(* IEC 61131-3 sources: daoli-st-library/DL_MathData (part 19) *)

(* ---- FC_DL_MeanAbsDevCalc.st ---- *)
(*
  ==================================================================
  组件名 Component  : FC_DL_MeanAbsDevCalc
  分类   Category   : DL_MathData
  前缀   Naming     : FC_DL_ ｜ b/n/u/f/t/e/st 类型前缀制（R265）
  复杂度 Complexity  : 低
  版本   Version    : 1.0.0
  功能   Purpose    : 均值绝对偏差 MAD-mean = mean(|xᵢ − mean|)，两遍法。
  来源   Source     : self-std（公开统计语义自研）
  平台   Platform   : 纯 IEC 61131-3（FOR / 四则 / ABS），三平台通用
  分工声明 Split     : 与 FC_DL_MedianAbsDev（中位数域属主）分工——后者以中位数
                      为中心（对离群点稳健）；本件以均值为中心（R216 双向互引）。
  作者   Author     : 道莅代码库 · PLC 编程专家（R61）
  归属 Ownership     : 本件无 TYPE 声明；引用件类型全部 IEC 标准原生。
  ------------------------------------------------------------------
  边界 Boundary     :
                      一 nCount < 1 置信息级码不计算（nCount = 0 无均值可言）；
                      二 计数 > 256 钳位续算置信息级；
                      三 元素非有限逐个点名判故障拒绝（R272 全量）；
                      四 均值非有限传播闸：均值算出后复检，非有限同判故障；
                      五 除子 nUse 已证 ≥ 1（域闸下界），无除零风险；
                      六 结果复检兜底同拍置 eErr + bError + bValid 三件套（R258）；
                      七 只读入参数组，不改调用方数据；无状态纯函数（R254）。
  错误码   Codes    :
    16#0001_063C【信息级】计数越域已钳位（<1 早退，>256 钳位续算）
    16#0001_063D【故障级】元素或均值非有限，拒绝出值
  验收   Acceptance :
    算法已证（脚本）：未跑 ｜ 编译器已证（三平台）：未跑
    V1 值 1/2/3 → mean=2、MAD-mean=2/3；V2 值 5/5/5 → 0
    V3 nCount=0 → 码 063C、bValid=FALSE；V4 含 NaN → 码 063D、bError=TRUE
  修订记录 Revision  :
    2026-11-21  v1.0.0  R61 首版（批 2 · 序号 7）
  ==================================================================
*)
FUNCTION FC_DL_MeanAbsDevCalc : BOOL
VAR_IN_OUT
    afValues : ARRAY[0..255] OF LREAL; // 数值序列 [工程单位]，只读 / the value series, read only
END_VAR
VAR_INPUT
    nCount : DINT; // 序列个数 [个]，合法域 1..256 / the count, legal from one to two hundred fifty six
END_VAR
VAR_OUTPUT
    fMad   : LREAL; // 均值绝对偏差 [工程单位] / the mean absolute deviation
    fMean  : LREAL; // 序列均值 [工程单位] / the series mean
    bValid : BOOL;  // 结果可用标志 [-] / the result usable flag
    eErr   : UDINT; // 错误码，0 = 正常 / the error code, zero is ok
    bError : BOOL;  // 错误标志，故障级码置位（R45 配对）/ the error flag
END_VAR
VAR
    k     : DINT;  // 遍历索引 [下标] / the traversal index
    nUse  : DINT;  // 钳位后的个数 [个] / the clamped count
    fSum  : LREAL; // 一遍和累加器 [工程单位] / the first pass sum accumulator
    fDev  : LREAL; // 二遍偏差累加器 [工程单位] / the second pass deviation accumulator
END_VAR
VAR CONSTANT
    DL_MAD_NMAX : DINT := 256; // 序列容量上界 [个]，与数组容量一致 / the capacity aligned with the array
END_VAR

// 段 1｜返回值与错误状态预置安全值 + 局部量显式预置（R45 / R254）/ segment 1, the preset
FC_DL_MeanAbsDevCalc := FALSE; // 返回值预置假 / preset the return false
fMad := 0.0; // 偏差预置零 / preset the deviation zero
fMean := 0.0; // 均值预置零 / preset the mean zero
bValid := FALSE; // 有效标志预置假 / preset the validity false
eErr := 16#0000_0000; // 错误码预置正常 / preset the code to ok
bError := FALSE; // 错误标志预置假 / preset the error flag false
nUse := 0; // 个数预置零 / preset the count zero
fSum := 0.0; // 一遍和预置零 / preset the sum zero
fDev := 0.0; // 二遍偏差预置零 / preset the deviation accumulator zero

// 段 2｜计数域闸（<1 早退，>256 钳位，边界一二）/ segment 2, the count gate
IF nCount < 1 THEN // 空序列无均值（边界一）/ an empty series has no mean
    eErr := 16#0001_063C; // 信息级：计数越域已钳位（信息级不置 bError）/ informational, the count clamped
    RETURN; // 早退 / early return
END_IF
nUse := nCount; // 域内接管 / take the count
IF nUse > DL_MAD_NMAX THEN // 超容量（边界二）/ above the capacity
    nUse := DL_MAD_NMAX; // 钳到容量 / clamp to the capacity
    eErr := 16#0001_063C; // 信息级：计数越域已钳位 / informational, the count clamped
END_IF

// 段 3｜一遍求和 + 元素非有限逐个点名（R272，边界三）/ segment 3, the first pass sum with the element wise gate
FOR k := 0 TO nUse - 1 DO // 有界遍历 / the bounded traversal
    IF (afValues[k] <> afValues[k]) OR ((afValues[k] - afValues[k]) <> (afValues[k] - afValues[k])) THEN // 元素非有限 / the element is not finite
        eErr := 16#0001_063D; // 故障级：元素非有限 / fault grade, a non finite element
        bError := TRUE; // 置错误标志（R45 配对）/ raise the error flag
        RETURN; // 早退 / early return
    END_IF
    fSum := fSum + afValues[k]; // 求和累加 / accumulate the sum
END_FOR
fMean := fSum / DINT_TO_LREAL(nUse); // 均值（除子已证 ≥ 1，边界五）/ the mean with a proven divisor
IF (fMean <> fMean) OR ((fMean - fMean) <> (fMean - fMean)) THEN // 均值非有限传播闸（边界四）/ the mean finiteness gate
    eErr := 16#0001_063D; // 故障级：均值非有限 / fault grade, a non finite mean
    bError := TRUE; // 置错误标志（R45 配对）/ raise the error flag
    RETURN; // 早退 / early return
END_IF

// 段 4｜二遍偏差累加（均值已证有限）/ segment 4, the second pass deviation accumulation
FOR k := 0 TO nUse - 1 DO // 有界遍历 / the bounded traversal
    fDev := fDev + ABS(afValues[k] - fMean); // 绝对偏差累加 / accumulate the absolute deviation
END_FOR
fMad := fDev / DINT_TO_LREAL(nUse); // 偏差均值（除子 nUse 已证 ≥ 1，同段 3 口径）/ the deviation mean with the proven divisor

// 段 5｜结果复检兜底（非有限同拍三件套，边界六）/ segment 5, the result recheck
IF (fMad <> fMad) OR ((fMad - fMad) <> (fMad - fMad)) THEN // 结果非有限 / the result is not finite
    fMad := 0.0; // 兜底安全值 / the bottom line safe value
    eErr := 16#0001_063D; // 故障级：结果非有限 / fault grade, the non finite result
    bError := TRUE; // 置错误标志（R45 配对）/ raise the error flag
    bValid := FALSE; // 结果不可用 / the result void
    RETURN; // 早退 / early return
END_IF
bValid := TRUE; // 结果可用 / the result is usable
FC_DL_MeanAbsDevCalc := TRUE; // 返回成功 / return success
END_FUNCTION

(* ---- FC_DL_MedianAbsDev.st ---- *)
(*==============================================================================
 * 组件名称 (Component)  : FC_DL_MedianAbsDev
 * 所属子库 (Sublibrary) : DL_MathData
 * 当前版本 (Version)    : 1.0.0
 * 兼容性   (Platform)   : CODESYS 3.5+ / TwinCAT 3 / 汇川 InoProShop / 施耐德 Machine Expert
 *                         仅用 FOR 循环、赋值与 ABS，无任何厂商内建函数（连排序库都不用）
 * 功能描述 (Function)   : 中位绝对偏差 MAD（Median Absolute Deviation），鲁棒离散度指标。
 *                           步骤：① 取前 nCount 个样本复制到本地缓冲（不改调用方数组）；
 *                                 ② 插入排序求中位数 fMedian；
 *                                 ③ 各样本减中位数取绝对值，再次插入排序求中位数 fMad。
 *                         返回 fMad。MAD 对离群点不敏感（崩溃点 50%），在传感器脏数据、
 *                         偶发尖峰场景下比标准差可靠：一个 10 倍离群点能把标准差抬高数倍，
 *                         而 MAD 几乎不变。
 *                         小样本策略：nCount < 3 → 无稳健意义，bValid=FALSE、返回 0；
 *                         nCount > 16 → 钳到 16（缓冲上界），bClamped=TRUE，结果按前 16 个算。
 *                         偶数样本的中位数取中间两数的算术平均（IEC 惯例，写死在此）。
 * 无状态边界 (Stateless): **本 FC 零内部状态**——本地缓冲 afWork / afDev 均为 VAR 临时量，
 *                         每次调用重新填装；IEC 61131-3 的 FC 本就不允许持有静态变量，本件遵守。
 *                         因此同一组样本重复调用结果完全一致，可重入、可并发、可放在任意 POU。
 *                         调用方若需"跨窗统计"，请自行保存样本数组，而不是期望 FC 记住上次数据。
 * 接口     (Interface)  : 入 afSample 样本数组（VAR_IN_OUT，本件只读，按 nCount 截取）、
 *                         nCount 有效样本数（1..16）；出 fMedian 中位数、fMad 中位绝对偏差、
 *                         bValid 结果有效（nCount >= 3）、bClamped 样本数被钳到 16。
 * 边界     (Boundary)   : ① 样本数下限：nCount < 3 无稳健离散意义 → bValid=FALSE、fMedian/fMad 置 0
 *                         （**0 不是"无离散"的断言**，调用方须查 bValid）；
 *                         ② 样本数上限：nCount > 16 → 钳到 16 并置 bClamped（绝不越 ARRAY 上界）；
 *                         ③ nCount <= 0 → bValid=FALSE、返回 0（防 nCount−1 为负导致的循环越界）；
 *                         ④ 非有限样本（NaN/Inf）会让排序结果失去意义：本件**不静默吞掉**，
 *                         检出即 bNonFin=TRUE、bValid=FALSE、返回 0（宁可不报，不可乱报）；
 *                         ⑤ 插入排序 O(n²)，n<=16 时最坏 256 次比较/两轮，代价可接受且无递归。
 * 依赖     (Depends)    : 无 DL_ 内部依赖；无标准库功能块依赖
 * 来源标签 (Source Tag) : T2-1 ◐（MAD 为公开经典鲁棒统计量，Hampel 1974；插入排序为教科书算法；
 *                         ST 实现为道莅自研，零代码行复制）
 * 码表     (Codes)      : 本件不占用任何全局数字码位。异常出口为 BOOL（bValid / bClamped / bNonFin）；
 *                         数字码位待主控收口阶段统一派号。
 * 红线自检 (Redline)    : R1 ✓ 零 GVL/VAR_EXTERNAL ｜ R2 ✓ 零 %I/%Q/%M ｜ R3 ✓ 纯 IEC 61131-3
 *                         R4 ✓ 数组边界钳位 + 循环上界由钳位量派生 + 非有限闸
 *                         R5 ✓ 声明逐行同行双语注释 ｜ R6 N/A（无状态机）
 *                         R7 N/A（无实例调用）
 * 修订历史 (Revision)   : 2026-11-19  v1.0.0  R46 首版（批次 3 · 序号 15）
 *==============================================================================*)
FUNCTION FC_DL_MedianAbsDev : REAL
VAR_IN_OUT
    afSample : ARRAY[0..15] OF REAL;    // 样本数组（本件只读，按 nCount 截取） [工程单位] / Sample array, read-only here, sliced by nCount
END_VAR
VAR_INPUT
    nCount : INT := 3;                  // 有效样本数，域 1..16（>16 被钳位） [个] / Valid sample count, 1..16, clamped above
END_VAR
VAR_OUTPUT
    fMedian  : REAL;                    // 样本中位数 [工程单位] / Sample median [engineering unit]
    bValid   : BOOL;                    // 结果有效（3 <= 有效样本数 <= 16） [-] / Result valid
    bClamped : BOOL;                    // 样本数被钳到 16 [-] / Sample count clamped to 16
    bNonFin  : BOOL;                    // 样本中存在 NaN/Inf，结果不可信 [-] / A non-finite sample was found
END_VAR
VAR
    afWork : ARRAY[0..15] OF REAL;      // 工作副本（排序用，不动调用方数组） [工程单位] / Working copy for sorting
    afDev  : ARRAY[0..15] OF REAL;      // 绝对偏差数组（排序用） [工程单位] / Absolute-deviation array for sorting
    nUse   : INT;                       // 实际参与计算的样本数（钳位后） [个] / Actual sample count after clamping
    i      : INT;                       // 外层遍历索引 / Outer loop index
    j      : INT;                       // 插入排序内层索引 / Inner index for the insertion sort
    fKey   : REAL;                      // 插入排序暂存键 [工程单位] / Key kept while inserting
    fLo    : REAL;                      // 偶数样本时中位数取中间两值之一 [工程单位] / One of the two middle values
    fHi    : REAL;                      // 偶数样本时中位数取中间两值之另一 [工程单位] / The other middle value
    nMidi  : INT;                       // 中位数取位下标（下中位） [个] / Lower middle index
END_VAR
VAR CONSTANT
    DL_MAD_MAXN : INT := 16;            // 样本容量（与 ARRAY 上界一致） [个] / Sample capacity matching the array bounds
    DL_MAD_MINN : INT := 3;             // 稳健统计所需最少样本数 [个] / Minimum sample count for robust statistics
END_VAR

(* —— 段 1：出口初始化（任何路径下返回值确定） —— *)
FC_DL_MedianAbsDev := 0.0;      // 缺省返回 0，须配 bValid 才可用 / Default 0, meaningful only with bValid
fMedian  := 0.0;                // 中位数清零 / Median cleared
bValid   := FALSE;              // 先假定无效 / Assume invalid
bClamped := FALSE;              // 钳位标志清零 / Clamp flag cleared
bNonFin  := FALSE;              // 非有限标志清零 / Non-finite flag cleared

(* —— 段 2：样本数钳位（先钳后循环，循环上界全部由 nUse 派生） —— *)
IF nCount <= 0 THEN
    RETURN;                     // 无样本：直接返回哨兵 0 / No samples: return the sentinel
END_IF
nUse := nCount;                 // 取请求样本数 / Take the requested count
IF nUse > DL_MAD_MAXN THEN
    nUse := DL_MAD_MAXN;        // 上界钳到容量 / Clamp to capacity
    bClamped := TRUE;           // 标记被钳 / Mark the clamp
END_IF

(* —— 段 3：复制到本地缓冲 + 非有限闸（NaN/Inf 会让排序失去意义，检出即拒算） —— *)
FOR i := 0 TO nUse - 1 DO
    afWork[i] := afSample[i];                               // 复制样本，不改调用方数组 / Copy, never modify the caller array
    IF (afWork[i] <> afWork[i]) OR ((afWork[i] - afWork[i]) <> (afWork[i] - afWork[i])) THEN
        bNonFin := TRUE;                                    // NaN 自反判 或 Inf 判（Inf−Inf 得 NaN） / NaN or Inf detected
    END_IF
END_FOR
IF bNonFin THEN
    RETURN;                     // 拒算：bValid 仍为假，返回 0 / Refuse: bValid stays false, 0 returned
END_IF

(* —— 段 4：插入排序（升序），小样本下比快排更省代码且无递归 —— *)
FOR i := 1 TO nUse - 1 DO
    fKey := afWork[i];                                      // 取出待插入键 / Take the key to insert
    j := i - 1;                                             // 从上一元素起向前扫 / Start scanning backwards
    WHILE (j >= 0) AND (afWork[j] > fKey) DO
        afWork[j + 1] := afWork[j];                         // 元素后移腾位 / Shift the element up
        j := j - 1;                                         // 索引前移（j 可到 −1，循环条件已含下界） / Step back, the loop condition covers -1
    END_WHILE
    afWork[j + 1] := fKey;                                  // 插入到位 / Insert at its place
END_FOR

(* —— 段 5：中位数（偶数样本取中间两值平均，写死口径） —— *)
nMidi := nUse / 2;                                          // 下中位下标（整除，nUse>=3 时 >=1） / Lower middle index
IF (nUse MOD 2) = 0 THEN
    fLo := afWork[nMidi - 1];                               // 中间左值 / Left middle value
    fHi := afWork[nMidi];                                   // 中间右值 / Right middle value
    fMedian := (fLo + fHi) * 0.5;                           // 偶数样本：算术平均 / Even count: arithmetic mean
ELSE
    fMedian := afWork[nMidi];                               // 奇数样本：正中值 / Odd count: the exact middle
END_IF

(* —— 段 6：绝对偏差数组 + 再次插入排序 —— *)
FOR i := 0 TO nUse - 1 DO
    afDev[i] := ABS(afWork[i] - fMedian);                   // 各样本到中位数的绝对距离 / Absolute distance to the median
END_FOR
FOR i := 1 TO nUse - 1 DO
    fKey := afDev[i];                                       // 取出待插入键 / Take the key
    j := i - 1;                                             // 从上一元素起向前扫 / Scan backwards
    WHILE (j >= 0) AND (afDev[j] > fKey) DO
        afDev[j + 1] := afDev[j];                           // 元素后移腾位 / Shift up
        j := j - 1;                                         // 索引前移 / Step back
    END_WHILE
    afDev[j + 1] := fKey;                                   // 插入到位 / Insert
END_FOR

(* —— 段 7：MAD 中位数 + 有效性判定（nUse >= 3 才算稳健） —— *)
nMidi := nUse / 2;                                          // 偏差数组的下中位下标 / Lower middle index of the deviations
IF (nUse MOD 2) = 0 THEN
    fLo := afDev[nMidi - 1];                                // 中间左值 / Left middle
    fHi := afDev[nMidi];                                    // 中间右值 / Right middle
    FC_DL_MedianAbsDev := (fLo + fHi) * 0.5;                // 偶数：平均 / Even: mean
ELSE
    FC_DL_MedianAbsDev := afDev[nMidi];                     // 奇数：正中值 / Odd: exact middle
END_IF
IF nUse >= DL_MAD_MINN THEN
    bValid := TRUE;                                         // 样本足够，结果有效 / Enough samples, result valid
ELSE
    bValid := FALSE;                                        // 样本过少，结果不宣称（返回值为 0） / Too few samples, nothing claimed
    FC_DL_MedianAbsDev := 0.0;                              // 明确置 0，避免半算值外溢 / Zero it explicitly
END_IF

END_FUNCTION

(* ---- FC_DL_MinEx.st ---- *)
(*
    FC_DL_MinEx —— 双值取小泛型防御包装（REAL 域）
    ------------------------------------------------------------------
    分类      : DL_MathData / MinMax
    前缀      : FC_DL_
    版本      : 1.0.0
    溯源      : IEC 61131-3 标准语义的道莅防御性实现
                （内部委托平台内建函数，外围统一错误码/钳位/双语文档；
                  未复制任何闭源厂商源码，参考实现仅限 MIT/Apache 许可）
    平台      : 纯 IEC 61131-3，CODESYS / TwinCAT / InoProShop 通用
    作者      : 道莅代码库 · PLC编程专家（R16）
    ------------------------------------------------------------------
    功能说明  : 双值取小：fA < fB 时返回 fA，否则返回 fB，比较运算委托
                `<` 运算符（IEC MIN 语义），不重实现任何数学内核；
                任一输入非有限（NaN 或 ±INF）判为故障级 16#0001_02B5，
                返回 0.0 且 bValid=FALSE（非有限值参与比较语义未定义，一律拦截）；
                钳位方向：无钳位（域内值直接比较输出，异常值故障拦截）；
                ±INF 采用平台安全幅值比较判定（阈值高于 REAL 最大有限值 3.402823E38），NaN 用自不等判定；
                信息级码位全部预留禁用（本组件无信息级路径）。
    错误码    : 16#0001_02B5 任一输入非有限（NaN 或 ±INF）——故障级，返回 0.0
                16#0001_01DA 预留禁用（信息级，不得挪用）
                16#0001_01DB 预留禁用（信息级，不得挪用）
                16#0001_02B6 预留禁用（故障级，不得挪用）
                16#0001_02B7 预留禁用（故障级，不得挪用）
    状态机    : R6 标注 N/A —— 本组件为纯函数无顺序状态机，无 CASE 可写，非法状态不可能出现，故以本节说明替代 ELSE 兜底
    修订记录  : 2026-11-16 v1.0.0 首次入库（R16）
*)
FUNCTION FC_DL_MinEx : REAL
VAR_INPUT
    fA : REAL; // 比较值 A [无量纲] / compare value A
    fB : REAL; // 比较值 B [无量纲] / compare value B
END_VAR
VAR_OUTPUT
    eErr   : UDINT; // 错误码，0=正常 / error id, 0=ok
    bError : BOOL;  // 是否出错，eErr 非 0 时为 TRUE / error flag, TRUE when eErr is nonzero
    bValid : BOOL;  // 输出是否有效可用 / output valid flag
END_VAR
VAR CONSTANT
    DL_REAL_INF_GUARD : LREAL := 4.0E38; // REAL 域 ±INF 判定阈值，高于 REAL 最大有限值 3.402823E38 [无量纲] / REAL +/-INF guard above max finite REAL 3.402823E38
END_VAR
VAR
    bBad : BOOL; // 任一输入非有限判定结果 / non-finite detection result of either input
END_VAR

// 段 1｜返回值与错误状态预置 / segment 1, preset return value and error status
FC_DL_MinEx := 0.0; // 故障缺省返回 0 [无量纲] / fault default returns 0
eErr   := 0;     // 预置无错误 / preset no error
bError := FALSE; // 预置无故障 / preset no fault
bValid := FALSE; // 预置无效，通过防御闸后置位 / preset invalid, set TRUE after guard passes

// 段 2｜非有限防御闸（末段：域内主体计算跟随） / segment 2, non-finite guard (final: in-domain main calculation follows)
bBad := (fA <> fA) OR (fA > DL_REAL_INF_GUARD) OR (fA < -DL_REAL_INF_GUARD)
     OR (fB <> fB) OR (fB > DL_REAL_INF_GUARD) OR (fB < -DL_REAL_INF_GUARD); // 双输入非有限判定（NaN 自不等 + 安全幅值判 ±INF） [无量纲] / both inputs non-finite check (NaN by self-inequality, +/-INF by safe magnitude)
IF bBad THEN
    FC_DL_MinEx := 0.0;       // 故障级返回 0 [无量纲] / fault level returns 0
    eErr   := 16#0001_02B5;   // 非有限输入故障码 / non-finite input fault id
    bError := TRUE;           // 置故障标志 / set fault flag
    bValid := FALSE;          // 输出无效 / output invalid
    RETURN;                   // 立即返回 / immediate return
END_IF

// 段 3｜域内取小主体计算 / segment 3, in-domain minimum main calculation
IF fA < fB THEN
    FC_DL_MinEx := fA; // A 较小，输出 A / A is smaller, output A
ELSE
    FC_DL_MinEx := fB; // B 较小或相等，输出 B（相等时二者同值） / B is smaller or equal, output B (identical when equal)
END_IF
bValid := TRUE; // 域内输出有效可用 / in-domain output is valid
END_FUNCTION

(* ---- FC_DL_MinNanEx.st ---- *)
(*
    FC_DL_MinNanEx —— 三输入取小内建防御包装（LREAL 域）
    ------------------------------------------------------------------
    分类      : DL_MathData / MinMax
    前缀      : FC_DL_
    版本      : 1.0.0
    溯源      : IEC 61131-3 标准语义的道莅防御性实现
                （内部委托平台内建函数 MIN，外围统一错误码/钳位/双语文档；
                  未复制任何闭源厂商源码，参考实现仅限 MIT/Apache 许可）
    平台      : 纯 IEC 61131-3，CODESYS / TwinCAT / InoProShop 通用
    作者      : 道莅代码库 · PLC编程专家（R40）
    ------------------------------------------------------------------
    功能说明  : 三输入取小：返回 fA、fB、fC 中的最小值，比较内核委托平台
                内建 MIN，不重实现任何数学内核；
                四段式口径（R45①）：返回值与错误码预置安全值 → 非有限域闸命中
                不调内建直接 RETURN → 域内委托内建 MIN → 结果非有限复检兜底；
                任一输入非有限判为故障级 16#0001_03CA，返回 0.0 且 bValid=FALSE
                （NaN 参与 MIN 比较在三平台传播行为不一致，一律拦截）；
                非有限判定口径（R15）：NaN 用自不等 f <> f 判定；±Inf 用
                (f − f) <> (f − f) 差值自减判定（有限值差恒为 0，无穷处产 NaN），
                禁用近似幅值阈值——LREAL 最大有限值 1.7976931348623157E308 之上
                无可表常量，近似阈值会在近似带内制造假阳性。
    错误码    : 16#0001_03CA 任一输入非有限（NaN 或 ±Inf）——故障级，返回 0.0
    状态机    : R6 标注 N/A —— 本组件为纯函数无顺序状态机，无 CASE 可写，
                非法状态不可能出现，故以本节说明替代 ELSE 兜底
    修订记录  : 2026-11-19 v1.0.0 首次入库（R40 · 批 1 · T0 快车道）
*)
FUNCTION FC_DL_MinNanEx : LREAL
VAR_INPUT
    fA : LREAL; // 候选值一 [无量纲] ｜ first candidate value
    fB : LREAL; // 候选值二 [无量纲] ｜ second candidate value
    fC : LREAL; // 候选值三 [无量纲] ｜ third candidate value
END_VAR
VAR_OUTPUT
    eErr   : UDINT; // 错误码，0=正常，16#0001_03XX=故障级 ｜ error id, 0=ok, 16#0001_03XX=fault level
    bError : BOOL;  // 是否出错，eErr 落故障级时为 TRUE ｜ fault flag, TRUE when eErr is fault level
    bValid : BOOL;  // 输出是否有效可用 ｜ output valid flag
END_VAR
VAR
    bBad : BOOL;  // 三输入非有限判定结果（NaN 或 ±Inf）｜ non-finite detection result of the three inputs
    fOut : LREAL; // 内建 MIN 结果暂存，供出口复检 ｜ staging of the MIN result for exit recheck
END_VAR

// 段 1｜返回值与错误状态预置 ｜ segment 1, preset return value and error status
FC_DL_MinNanEx := 0.0; // 故障缺省返回 0 [无量纲] ｜ fault default returns 0
eErr   := 0;     // 预置无错误 ｜ preset no error
bError := FALSE; // 预置无故障 ｜ preset no fault
bValid := FALSE; // 预置无效，通过防御闸后置位 ｜ preset invalid, set TRUE after guard passes
fOut   := 0.0;   // 暂存清零 ｜ clear the staging value

// 段 2｜三输入非有限防御闸（命中不调内建，早退） ｜ segment 2, non-finite guard of the three inputs (early return, no built-in call)
bBad := (fA <> fA) OR ((fA - fA) <> (fA - fA))
     OR (fB <> fB) OR ((fB - fB) <> (fB - fB))
     OR (fC <> fC) OR ((fC - fC) <> (fC - fC)); // 三输入非有限判定：NaN 自不等 + 差值自减判 ±Inf [无量纲] ｜ non-finite check: NaN by self-inequality, +/-Inf by self-subtraction
IF bBad THEN
    FC_DL_MinNanEx := 0.0;  // 故障级返回 0 [无量纲] ｜ fault level returns 0
    eErr   := 16#0001_03CA; // 非有限输入故障码 ｜ non-finite input fault id
    bError := TRUE;         // 置故障标志（R45 配对）｜ raise the fault flag (R45 pairing)
    bValid := FALSE;        // 输出无效 ｜ output invalid
    RETURN;                 // 早退，不调内建 ｜ early return, no built-in call
END_IF

// 段 3｜域内委托内建 MIN 内核 ｜ segment 3, delegate to the built-in MIN kernel in domain
fOut := MIN(fA, fB, fC); // 三输入取小委托内建 [无量纲] ｜ three-input minimum delegated to the built-in

// 段 4｜结果复检兜底（理论不可达：有限值的 MIN 恒有限） ｜ segment 4, exit recheck (unreachable: MIN of finite values is finite)
IF (fOut <> fOut) OR ((fOut - fOut) <> (fOut - fOut)) THEN
    FC_DL_MinNanEx := 0.0;  // 复检失败按非有限处置 [无量纲] ｜ recheck failure treated as non-finite
    eErr   := 16#0001_03CA; // 复用非有限输入码（同因同码，不新占码位）｜ reuse the non-finite code (same cause, no new code)
    bError := TRUE;         // 置故障标志 ｜ raise the fault flag
    bValid := FALSE;        // 输出无效 ｜ output invalid
    RETURN;                 // 早退 ｜ early return
END_IF

// 段 5｜出口装配 ｜ segment 5, exit assembly
FC_DL_MinNanEx := fOut; // 取小结果直通 ｜ minimum result pass-through
bError := FALSE;        // 正常出口不置故障 ｜ normal exit raises no fault
bValid := TRUE;         // 输出有效可用 ｜ output valid
END_FUNCTION

(* ---- FC_DL_ModLrealSafe.st ---- *)
(*==============================================================================
 * 组件名称 (Component)  : FC_DL_ModLrealSafe
 * 所属子库 (Sublibrary) : DL_MathData
 * 归属目录 (Directory)  : C:\Library\DL_MathData
 * 当前版本 (Version)    : 1.0.0
 * 分类/来源标签         : 函数（FUNCTION）· 纯函数 · LREAL 安全取模
 *                         iec-std-wrapper / math-safe
 * 兼容性   (Platform)   : CODESYS 3.5 / TwinCAT 3 / 汇川 InoProShop / 施耐德
 *                         Machine Expert；仅用 IEC 标准算术与 TRUNC 语义
 * 溯源声明 (Provenance) : IEC 61131-3 标准语义的道莅防御性实现——内部委托平台标准库语义，
 *                         外围统一错误码 / 钳位 / 双语注释，严禁重实现数学内核。
 * 功能一句话 (Summary)  : LREAL 安全取模：除零与绝对小除数双闸、输入非有限闸、
 *                       结果非有限闸四道防线，防 NaN 沿数据链扩散。
 *
 * 功能描述 (Function)   : 四闸顺序：① 输入非有限闸（NaN 自反判据、Inf 实数上限
 *                         判据）；② 除零闸（除数绝对值小于 fEps 视为零，防浮点
 *                         下溢假非零）；③ 商域闸（商绝对值超过 DL_MAXQ 时 TRUNC
 *                         会溢出整数域，直接拒绝）；④ 结果非有限闸。合法路径用
 *                         标准 fA - fB * TRUNC(fA / fB) 表达式实现取模，零被除数
 *                         以信息级告知恒等余数零。
 * 与既有件边界 (Boundary): 与 FC_DL_DivLrealSafe 组成除/模对；本件不做浮点取整
 *                         方向选择（floor/ceil 变体归后续件），固定向零截断。
 * 码位说明 (Codes)      : 信息 16#0002_3050 零被除数恒等（余数为零）
 *                         故障 16#0002_3051 除数无效（零或绝对值小于 fEps）
 *                         故障 16#0002_3052 输入非有限（NaN 或 Inf）
 *                         故障 16#0002_3053 结果域外（商超界或结果非有限）
 *                         段 16#02_3_50~53 首槽信息级、次槽起故障级。
 * 依赖说明 (Depends)    : 无 DL_ 内部依赖；仅 IEC 标准算术 / ABS / TRUNC。
 * 红线自检 (Redline)    : 零全局依赖 ｜ 零 VAR_EXTERNAL ｜ 零 %I/%Q ｜ 纯 IEC 标准库
 *                         浮点比较全部带 fEps 容差 ｜ NaN/Inf 用精确判据
 *                         除法前强制判零 ｜ 全变量双语同行注释 ｜ 无定时器实例
 * 修订历史 (Revision)   : 2026-11-18  v1.0.0  首版入库（R32 · 批 2）
 *============================================================================*)

FUNCTION FC_DL_ModLrealSafe : BOOL
VAR_INPUT
    fA    : LREAL;                  // 被除数 [实数域] / Dividend
    fB    : LREAL;                  // 除数 [实数域]，绝对值小于 fEps 视为零 / Divisor, near-zero by fEps
    fEps  : LREAL := 1.0E-12;       // 判零容差 [实数域] / Zero tolerance
END_VAR
VAR_OUTPUT
    fRem    : LREAL;                // 余数 [实数域]，故障路径为哨兵零 / Remainder, sentinel zero on fault
    bError  : BOOL;                 // 故障标志，与故障码 3051~3053 配对 / Fault flag paired with codes
    uErrorId: UDINT;                // 事件码，0 表示无事件 / Event code, zero means none
END_VAR
VAR
    fQ   : LREAL;   // 中间商 [实数域]，仅作域判定与截断 / Intermediate quotient
    uCode: UDINT;   // 码位暂存，出口单点写入 [码] / Code staging
END_VAR
VAR CONSTANT
    DL_MLS_MAXQ : LREAL := 1.0E9;   // 商绝对值上限 [实数域]，保 TRUNC 不溢出 DINT / Quotient cap, keeps TRUNC inside DINT
END_VAR

(* 段 1｜输出预置 / Pre-set *)
FC_DL_ModLrealSafe := FALSE;
fRem     := 0.0;
bError   := FALSE;
uErrorId := 16#0000_0000;
uCode    := 16#0000_0000;

(* 段 2｜输入非有限闸：NaN 自反判据、Inf 实数上限判据 / Non-finite input gate *)
IF (fA <> fA) OR (fB <> fB) OR (ABS(fA) > 1.0E308) OR (ABS(fB) > 1.0E308) THEN
    fRem    := 0.0;              // 哨兵零 / Sentinel zero
    bError  := TRUE;             // 故障级码配对置位 / Fault flag paired
    uErrorId := 16#0002_3052;    // 故障级：输入非有限 / Fault: non-finite input
    RETURN;
END_IF

(* 段 3｜除零闸：精确零与绝对小除数一并拦截，防浮点下溢假非零 / Zero gate: exact zero and near-zero together *)
IF ABS(fB) < fEps THEN
    fRem    := 0.0;              // 哨兵零 / Sentinel zero
    bError  := TRUE;             // 故障级码配对置位 / Fault flag paired
    uErrorId := 16#0002_3051;    // 故障级：除数无效 / Fault: invalid divisor
    RETURN;
END_IF

(* 段 4｜零被除数恒等：信息级告知 / Zero dividend identity *)
IF ABS(fA) < fEps THEN
    fRem    := 0.0;              // 恒等余数零 / Identity remainder zero
    uErrorId := 16#0002_3050;    // 信息级：零被除数 / Info: zero dividend
    FC_DL_ModLrealSafe := TRUE;
    RETURN;
END_IF

(* 段 5｜商域闸：商超界时 TRUNC 会溢出整数域，拒绝而不硬算 / Quotient domain gate: refuse before TRUNC could overflow *)
fQ := fA / fB;
IF ABS(fQ) > DL_MLS_MAXQ THEN
    fRem    := 0.0;              // 哨兵零 / Sentinel zero
    bError  := TRUE;             // 故障级码配对置位 / Fault flag paired
    uErrorId := 16#0002_3053;    // 故障级：结果域外 / Fault: result out of domain
    RETURN;
END_IF

(* 段 6｜合法路径：标准向零截断取模表达式 / Legal path: standard truncation-based modulo *)
fRem := fA - fB * TRUNC(fQ);     // fA 减 fB 乘整数商得余数 / Dividend minus divisor times truncated quotient

(* 段 7｜结果非有限闸（防御校验，正常路径不可达）/ Result non-finite gate, belt and braces *)
IF (fRem <> fRem) OR (ABS(fRem) > 1.0E308) THEN
    fRem    := 0.0;              // 哨兵零 / Sentinel zero
    bError  := TRUE;             // 故障级码配对置位 / Fault flag paired
    uErrorId := 16#0002_3053;    // 故障级：结果非有限 / Fault: non-finite result
    RETURN;
END_IF
uErrorId := uCode;               // 码位单点写入 / Single write point
FC_DL_ModLrealSafe := TRUE;
END_FUNCTION

(* ---- FC_DL_ModPos.st ---- *)
(*
    组件名称 : FC_DL_ModPos
    所属子库 : DL_MathData
    当前版本 : 1.0.0
    兼 容 性 : CODESYS V3.5+ / TwinCAT 3 / 汇川 InoProShop；仅依赖 Standard.library
    功能描述 : 恒正取模原子，返回恒非负余数 r ∈ [0, |m|-1]，消灭「负数取余」在三大平台上的符号歧义。
              取舍 ①：全文只允许一次 MOD —— 先按模数绝对值取余，再用「条件加法」把负余数搬回正域。
              禁二次取模（r := (v MOD m + m) MOD m），那是同一歧义的第二处实现，改一处必漏一处。
              取舍 ②：禁「先 ABS 再 MOD」。ABS(nValue) 在 nValue = DINT_MIN 处回绕成自身，会静默算错；
              本件只对模数取绝对值，并对 DINT_MIN 模数直接报故障。
              取舍 ③：模数为负时取绝对值后照算并发信息级提示 —— (-7) MOD (-3) 与 (-7) MOD 3 归一后同为 2，
              模数符号不影响数学结论，但调用方多半写错了，必须让它看得见而不是静默吞掉。
    开源溯源 : 原创实现。取模归一属 IEC 61131-3 MOD 运算符的防御性封装，无外部源码参考；；本件为 IEC 61131-3 标准语义的道莅防御性实现（原创实现，零外部源码复制）。
              码位、错误分级、下界哨兵策略与注释 100% 自有。
    本文件内含 : FUNCTION FC_DL_ModPos（单 POU，无配套类型）
    依 赖 : 无 DL_ 内部依赖；Standard.library: 无
    红线自检 : R1 ✓ 零全局变量与外部变量 ｜ R2 ✓ 零物理 IO 地址
              R3 ✓ 纯 IEC 61131-3 ｜ R4 ✓ 零模闸 + 下界闸 + 条件加法归一（无二次取模、无 ABS 单侧）
              R5 ✓ 全变量中英双语同行注释 ｜ R6 N/A 纯函数无顺序状态机，无 CASE 可写
              R7 N/A 无定时器、无沿检测实例 ｜ R8 ✓ 全部哨兵与下界常量化
    错误码   : 16#0001_0434 [信息级] 模数为负已取绝对值，结果照算，bError = FALSE，bValid = TRUE
               16#0001_0435 [信息级] 预留禁用（不得挪用）
               16#0001_036C [故障级] 模数为零，返回 0，bValid = FALSE
               16#0001_036D [故障级] 模数为 DINT 下界，取绝对值溢出，返回 0，bValid = FALSE
               16#0001_036E [故障级] 预留禁用（不得挪用）
    码位总账 : 16#0001_0434 用 / 16#0001_0435 预留 ｜ 16#0001_036C 用 / 16#0001_036D 用 / 16#0001_036E 预留
    遗留假设 : ① MOD 余数符号按 IEC 61131-3 取「与被除数同号」，本件的条件加法同时兼容「恒非负」与「同号」
              两种平台实现，故该假设失效也不改变结果 —— 此结论为推导，未在三平台逐一实测。
              ② 本件无内建转换链、无时间日期口径，编译门槛未见风险。
    修订历史 :
        2026-11-16  v1.0.0  首版，R21 批次 1 入库
*)
FUNCTION FC_DL_ModPos : DINT
VAR_INPUT
    nValue          : DINT;   // 被除数，全域 -2147483648~2147483647 [无量纲] / dividend, full DINT domain [dimensionless]
    nModulus        : DINT;   // 模数，必须 ≠ 0；为负时取绝对值后照算 [无量纲] / modulus, must not be zero, negative modulus is taken by absolute value [dimensionless]
END_VAR
VAR_OUTPUT
    eErr            : UDINT;  // 错误码，0=正常；16#0001_04XX 信息级 / 16#0001_03XX 故障级 / error id, 0=ok
    bError          : BOOL;   // 故障级标志，eErr 落 16#0001_03XX 时为 TRUE / fault flag, TRUE on fault-level eErr
    bValid          : BOOL;   // 返回值是否可用，FALSE 时调用方必须走故障分支 / output valid flag, the caller must branch when FALSE
END_VAR
VAR
    nModAbs         : DINT;   // 模数绝对值，进入取模前恒 > 0 [无量纲] / absolute modulus, always positive before the MOD [dimensionless]
    nRem            : DINT;   // 余数工作寄存器，出口前被搬入正域 [无量纲] / remainder working register, moved into the positive domain before exit [dimensionless]
END_VAR
VAR CONSTANT
    DL_DINT_ZERO    : DINT := 0;             // 零哨兵，避免裸 0 参与比较 [无量纲] / zero sentinel, no bare zero in comparisons [dimensionless]
    DL_DINT_MIN     : DINT := -2147483648;   // DINT 下界，取绝对值回绕，必须单独拦截 [无量纲] / DINT lower bound whose absolute value wraps around [dimensionless]
    DL_DINT_MIN_ABS : DINT := -2147483647;   // 可直接取绝对值的下界哨兵（−MAX−1 的邻值）[无量纲] / lowest value that can be negated safely [dimensionless]
    DL_ERR_NONE     : UDINT := 16#0000_0000; // 无故障 / no error
END_VAR

// 段 1｜返回值与错误状态预置（四段式第一段）/ segment 1, preset the return value and the error state
FC_DL_ModPos := DL_DINT_ZERO;   // 故障缺省返回 0 / fault default returns zero
eErr         := DL_ERR_NONE;    // 预置无错误 / preset no error
bError       := FALSE;          // 预置无故障 / preset no fault
bValid       := FALSE;          // 预置结果不可用，通过全部闸门后置 TRUE / preset unusable, set TRUE after every gate
nModAbs      := nModulus;       // 先按原值占位，符号归一后会覆盖 / provisional copy, overwritten by the sign normalisation

// 段 2｜模数零闸：零模一律不进 MOD / segment 2, zero modulus gate, never enter the MOD
IF nModulus = DL_DINT_ZERO THEN
    eErr   := 16#0001_036C;     // 模数为零（故障级）/ zero modulus, fault level
    bError := TRUE;             // 置故障标志 / raise the fault flag
    RETURN;                     // 返回 0，bValid 保持 FALSE / return zero, bValid stays FALSE
END_IF

// 段 3｜模数下界闸：DINT_MIN 取绝对值回绕成自身，必须拒算 / segment 3, lower bound gate, negating DINT_MIN wraps around
IF nModulus = DL_DINT_MIN THEN
    eErr   := 16#0001_036D;     // 模数下界不可表示其绝对值（故障级）/ modulus lower bound has no representable absolute value
    bError := TRUE;             // 置故障标志 / raise the fault flag
    RETURN;                     // 返回 0，bValid 保持 FALSE / return zero, bValid stays FALSE
END_IF

// 段 4｜模数符号归一：负模取绝对值，信息级提示，结果照算 / segment 4, negative modulus is normalised, info level only
IF nModulus < DL_DINT_ZERO THEN
    nModAbs := -nModulus;       // 下界已拦，取负结构性安全 / the lower bound is already rejected, so negation is structurally safe
    eErr    := 16#0001_0434;    // 模数为负已取绝对值（信息级，不置 bError）/ negative modulus normalised, info level, never sets bError
END_IF

// 段 5｜全文唯一一次 MOD，然后条件加法把负余数搬回正域 / segment 5, the single MOD followed by one conditional add
nRem := nValue MOD nModAbs;     // 余数与被除数同号，负域需归一 / the remainder follows the dividend sign and must be normalised
IF nRem < DL_DINT_ZERO THEN
    nRem := nRem + nModAbs;     // 加一次模数即落回 [0, |m|-1]，不做二次取模 / one addition lands in [0, |m|-1], no second MOD
END_IF

// 段 6｜出口：结果是真值，bValid 置 TRUE / segment 6, exit with a genuine value
FC_DL_ModPos := nRem;           // 输出归一后的非负余数 / publish the normalised non-negative remainder
bValid       := TRUE;           // 结果可用（信息级不影响可用性）/ the result is usable, info codes never block it
END_FUNCTION

(* ---- FC_DL_ModPosWrap.st ---- *)
(*
    FC_DL_ModPosWrap —— 取模正值回绕（负余数归正）
    ------------------------------------------------------------------
    组件名称  : FC_DL_ModPosWrap
    分类      : DL_MathData / IntegerArith
    前缀      : FC_DL_
    版本      : 1.0.0
    溯源      : 借鉴点 —— IEC 61131-3 第 3 版整数 MOD 运算符的标准语义
                （余数符号随被除数，即截断除法口径）；本件把该口径**归一到
                非负区间**，即数学意义上的「正模」语义，供环形缓冲下标、
                角度索引、多工位轮转相位等需要恒非负余数的场合使用。
                clean-room 声明 —— 零代码行复制，仅调用平台内建 MOD 运算符，
                外围的域闸 / 归正 / 码位 / 双语文档全部自有。
                许可证 —— 本件 MIT；标准文本仅作语义引用，不构成代码许可继承。
    平台      : 纯 IEC 61131-3，CODESYS 3.5 / TwinCAT 3 / InoProShop / Machine Expert 通用
    作者      : 道莅代码库 · PLC编程专家（R70 构建轮 · 批 1 · N1）
    ------------------------------------------------------------------
    功能说明  : 计算 liValue 对 liMod 的非负取模，结果恒落在 [0, |liMod|) 区间。
                与库内既有件的分工（防止重复实现）：
                  FC_DL_ModPos（DL_MathData）为 DINT 版同类语义；
                  本件为 LINT 64 位版，并把「负模数」也纳入契约：libs 内建 MOD
                  在模数为负时余数符号不可直接用，本件显式归一，故返回值区间
                  与模数符号无关。
                归正算法的双语义兼容性（关键设计）：内建 MOD 在截断除法口径下
                返回负余数，在部分平台的实现中也可能已返回非负余数。本件仅做
                一次条件补正 —— 余数 < 0 时按模数符号分别 +m 或 -m —— 对两种
                内建语义均得到同一正确结果，不依赖平台细节。
                溢出安全性（逐分支论证）：设 m = |liMod| > 0，内建余数 r 满足
                |r| < m。r < 0 且 liMod > 0 时取 r + liMod，落在 (0, m) 内；
                r < 0 且 liMod < 0 时取 r - liMod 即 r + m，落在 (0, m) 内；
                两条路径的结果绝对值均小于 2^63，不存在 LINT 溢出；
                模数为 LINT 下界时 m 不可直接取绝对值，故本件**不对模数取绝对值**，
                只按符号选择运算方向，从而绕开 |LINT_MIN| 不可表示的问题。
    错误码    : 16#0002_0101 模数为 0（除零禁入），返回 0 —— 故障级
                16#0002_0102 保留（LINT 下界模数无需特殊处理，见上论证）—— 未用
    码位总账  : 16#0002_0101 用 ｜ 16#0002_0102 保留未用
    状态机    : R6 N/A —— 纯函数无状态，无跨周期驻留，无 CASE 可写
    边界与披露: 一 无定时器 / 无边沿实例 / 无除法 / 无数组下标，周期安全规则 N/A；
                二 零全局变量、零 VAR_EXTERNAL、零物理地址，纯引脚契约；
                三 bNegAdjusted 仅在「内建余数为负并被补正」时为 TRUE，
                   供上层统计平台语义差异，不参与任何判据；
                四 模数为 0 时按契约返回 0 且置故障级码，bValid = FALSE，
                   调用方必须用 bValid 或 bError 门控返回值，不得直取。
    修订记录  : 2026-11-22 v1.0.0 首次入库（R70 构建轮 · 批 1 · N1）
*)
FUNCTION FC_DL_ModPosWrap : LINT
VAR_INPUT
    liValue : LINT;                        (* 被除数（可为负），[计数] / the dividend, may be negative *)
    liMod   : LINT;                        (* 模数（非零），[计数]，符号自动归一 / the modulus, non-zero, sign normalised *)
END_VAR
VAR_OUTPUT
    eErr         : UDINT;                  (* 错误码，0 = 正常 / the error id, 0 = ok *)
    bError       : BOOL;                   (* 故障标志，故障级码时 TRUE / the error flag, TRUE on fault level *)
    bValid       : BOOL;                   (* 返回值可用，故障级为 FALSE / the return usable, FALSE on fault level *)
    bNegAdjusted : BOOL;                   (* 内建余数为负且已补正，[标志] / the negative remainder was corrected *)
END_VAR

// 段 1｜返回值与状态预置（四段式第一段）/ segment 1, preset the return and the status
FC_DL_ModPosWrap := 0;                 // 故障缺省返回 0 / the fault default returns 0
eErr         := 0;                     // 预置无错误 / preset no error
bError       := FALSE;                 // 预置无故障 / preset no fault
bValid       := FALSE;                 // 预置不可用，过闸后置位 / preset unusable, set TRUE after the gates
bNegAdjusted := FALSE;                 // 预置未补正 / preset not corrected

// 段 2｜除零域闸：模数为 0 结构早退，绝不落除法内核 / segment 2, the zero modulus gate, structural early return
IF liMod = 0 THEN                      // 模数为零即除零，禁入 / a zero modulus means a division by zero
    eErr   := 16#0002_0101;            // 故障级：模数为 0 / fault level: the modulus is zero
    bError := TRUE;                    // R45 配对置故障标志 / paired with the code
    bValid := FALSE;                   // 返回值不可用 / the return is unusable
    RETURN;                            // 结构早退，内建 MOD 不被触碰 / structural exit, the MOD kernel is never touched
END_IF

// 段 3｜委托内建 MOD 内核（模数已证非零）/ segment 3, delegate to the built-in MOD kernel
FC_DL_ModPosWrap := liValue MOD liMod; // 内建取模，余数符号随平台口径 / the built-in remainder, sign per the platform

// 段 4｜负余数归正：按模数符号选择补正方向，避免对 LINT 下界取绝对值 / segment 4, normalise a negative remainder
IF FC_DL_ModPosWrap < 0 THEN           // 内建余数为负（截断除法口径）/ a negative remainder, the truncated convention
    bNegAdjusted := TRUE;              // 记录已补正 / record the correction
    IF liMod > 0 THEN                  // 正模数：加模数即入正域 / a positive modulus, add it
        FC_DL_ModPosWrap := FC_DL_ModPosWrap + liMod;   // 结果落 (0, m) / the result lands in (0, m)
    ELSE                               // 负模数：减模数即加 |m|（不取绝对值，避开 LINT_MIN）/ a negative modulus, subtract it
        FC_DL_ModPosWrap := FC_DL_ModPosWrap - liMod;   // 结果落 (0, |m|) / the result lands in (0, |m|)
    END_IF
END_IF

// 段 5｜出口状态：域内委托结果恒可用 / segment 5, the outlet status, an in-domain result is always usable
bError := FALSE;                       // 本路径无故障 / no fault on this path
bValid := TRUE;                        // 余数可用 / the remainder is usable
END_FUNCTION

(* ---- FC_DL_MoistureContentCalc.st ---- *)
// FC_DL_MoistureContentCalc v1.0.0
// 开源溯源：self-cleanroom / 公开公式（失重法含水率）
(*
  道莅工业代码库 | DL_MathData | FC_DL_MoistureContentCalc
  版本: 1.0.0 | 日期: 2026-11-23 | 轮次: R75
  功能: 失重法含水率计算：(湿重 - 干重) / 湿重 × 100%，湿重分母域闸 +
        干湿重序闸（干 > 湿 判测量矛盾）
  邻件关系: 与 ElectrolyteMoistureGuard（电解液含水防护联锁）相邻 ——
            差异点：防护件为阈值联锁动作，本件为纯计算件（无联锁输出），
            工业称重/烘干域通用
*)
FUNCTION FC_DL_MoistureContentCalc : REAL
VAR_INPUT
    fWetMassG : REAL := 0.0;    // 湿重 [g]，域 > 0 / Wet mass [g], domain > 0
    fDryMassG : REAL := 0.0;    // 干重 [g]，域 >= 0 且 <= 湿重 / Dry mass [g], domain >= 0 and <= wet
    fEps      : REAL := 1.0E-6; // 判零容差 [g] / Zero tolerance [g]
END_VAR
VAR_OUTPUT
    bValid    : BOOL;           // 结果有效回执 [-] / Result validity receipt
    uErrorId  : UDINT;          // 事件码，0 = 无事件；16#0002_2001 = 域外拒收 / Event code
END_VAR

// —— 段 0：全路径缺省 —— //
bValid   := FALSE;              // 有效回执预清 / Validity preset
uErrorId := 16#0000;            // 事件码预清 / Event code preset
FC_DL_MoistureContentCalc := 0.0;   // 返回值缺省零 / Return default zero

// —— 段 1：非有限闸 —— //
IF (fWetMassG <> fWetMassG) OR (fDryMassG <> fDryMassG)
   OR (ABS(fWetMassG) >= 3.0E38) OR (ABS(fDryMassG) >= 3.0E38) THEN
    uErrorId := 16#0002_2001;   // 输入非有限拒收（域闸码复用，R90 不加码）/ Non-finite reject
    RETURN;
END_IF

// —— 段 2：域闸（湿重正数 + 干湿序 + 负干重拒收） —— //
IF (fWetMassG < fEps) OR (fDryMassG < 0.0) OR (fDryMassG > fWetMassG) THEN
    uErrorId := 16#0002_2001;   // 信息级：湿重近零/干重为负/干重超湿重（测量矛盾）/ Info level: domain violation
    RETURN;                     // 不计算返回零 / Return zero without division
END_IF

// —— 段 3：主计算（分母已过闸） —— //
FC_DL_MoistureContentCalc := (fWetMassG - fDryMassG) / fWetMassG * 100.0;   // 含水率 [%] / Moisture content [%]
bValid := TRUE;                 // 有效回执 / Validity receipt
END_FUNCTION

(* ---- FC_DL_MolassesExhaustionCalc.st ---- *)
(*
  Component : FC_DL_MolassesExhaustionCalc
  Category  : DL_MathData
  Type      : FC
  Complexity: C1
  VERSION   : v1.0.0
  功能      : 废蜜纯度与糖分排出率核算：按糖膏纯度与废蜜纯度算糖分排出率（提净率）与随废蜜损失的糖分比例。
  开源溯源  : 道莅原创 clean-room 自研（无外部代码引用）｜License: MIT
  边界条件  : ① 糖膏纯度须 > 1e-9（为除子），否则返回哨兵 -1；
              ② 废蜜纯度高于糖膏纯度时排出率为负（数据异常），照实输出供诊断不钳位；
              ③ 两个纯度均须落在 0~100 % 理化可表区间。
*)
FUNCTION FC_DL_MolassesExhaustionCalc : REAL
VAR_INPUT
    fMassePurityPct   : REAL;   (* 糖膏（母液）纯度 [%] Massecuite purity *)
    fMolassesPurityPct: REAL;   (* 废蜜纯度 [%] Molasses purity *)
END_VAR
VAR_OUTPUT
    fExhaustPct : REAL;   (* 糖分排出率（提净率） [%] Exhaustion percent *)
    fLossPct    : REAL;   (* 随废蜜损失的糖分比例 [%] Sugar loss percent *)
    xValid      : BOOL;   (* 计算有效性标志 [-] Calculation valid flag *)
END_VAR
VAR CONSTANT
    DL_EPS      : REAL := 1.0E-9;   (* 除零判定容差 [无量纲] Divide-by-zero tolerance *)
    DL_PCT_BASE : REAL := 100.0;    (* 百分比基准 [%] Percent base *)
    DL_ZERO     : REAL := 0.0;      (* 零常量 [无量纲] Zero constant *)
END_VAR
(* 出口预置：三出口统一预置 *)
fExhaustPct := 0.0; fLossPct := 0.0; xValid := FALSE;
(* 非有限拦截：自反判 NaN，自身差值判 Inf *)
IF (fMassePurityPct <> fMassePurityPct) OR ((fMassePurityPct - fMassePurityPct) <> 0.0)
   OR (fMolassesPurityPct <> fMolassesPurityPct)
   OR ((fMolassesPurityPct - fMolassesPurityPct) <> 0.0) THEN
    FC_DL_MolassesExhaustionCalc := -1.0;  (* 哨兵 -1：输入非有限 / Sentinel -1 non-finite *)
    RETURN;
END_IF
(* 理化域闸：糖膏纯度为除子，两纯度须落在 0~100 % *)
IF (fMassePurityPct <= DL_EPS) OR (fMassePurityPct > DL_PCT_BASE)
   OR (fMolassesPurityPct < DL_ZERO) OR (fMolassesPurityPct > DL_PCT_BASE) THEN
    FC_DL_MolassesExhaustionCalc := -1.0;  (* 哨兵 -1：组态非法 / Sentinel -1 bad config *)
    RETURN;
END_IF
(* 糖分排出率：(糖膏纯度 - 废蜜纯度) / 糖膏纯度，除子已过域闸 *)
fExhaustPct := (fMassePurityPct - fMolassesPurityPct) / fMassePurityPct * DL_PCT_BASE;
(* 糖分损失比例：废蜜纯度占糖膏纯度的份额 *)
fLossPct := fMolassesPurityPct / fMassePurityPct * DL_PCT_BASE;
xValid := TRUE;                           (* 链路有效 / Chain valid *)
FC_DL_MolassesExhaustionCalc := fExhaustPct;  (* 返回排出率 [%] / Return exhaustion percent *)
END_FUNCTION

(* ---- FC_DL_MovingRangeCalc.st ---- *)
//==============================================================================
// 函数：FC_DL_MovingRangeCalc ｜ 中文名称：滑动极差（相邻样本差）原子计算
// 所属子库：DL_MathData ｜ 版本：v1.0.0 ｜ 日期：2026-11-23
// 兼容：CODESYS V3.5+ / TwinCAT 3 / 汇川 InoProShop / Machine Expert（纯标准库）
// 功能描述：SPC 判稳前置原子：MR = |x_i − x_(i−1)|，相邻两样本的极差。
//           无状态原子：本拍新样本与上一拍样本由调用方传入，本件不驻留
//           历史样本（滑动窗管理属上层 FB，职责边界见头注释）。
// 开源溯源 (Origin)：原创实现（t2-1-lgf-measurement 测量链语义深化，零外部
//           源码行，clean-room 独立编写）
// 公开接口清单：输入 fNewSample / fPrevSample；输出 fRange / bValid
// 单位表：fNewSample / fPrevSample / 返回值 [工程单位随调用方，差值不改单位]
// 输入契约：两样本须同一工程单位同一测点（跨测点差值无物理意义）；调用方
//           负责滑动窗历史驻留与回传节奏。
// 输出契约：返回值为极差（恒非负）；bValid = FALSE 拍返回哨兵 0.0，
//           调用方禁将哨兵值计入 SPC 控制图样本。
// 错误码表：纯函数无状态机码轨；无效输入经 bValid = FALSE 表达（哨兵返回
//           0.0），本件不占用 16#0001 段码位（邻件免让位）
// 状态机：N/A（纯函数，无状态，可重入）
// 边界行为：① 任一输入非有限（NaN 自反判 + 幅值上限判）→ bValid := FALSE、
//           哨兵 0.0 返回；② 极差恒非负（ABS 内建保证）；③ 无除法无域闸。
// 修订历史：v1.0.0 2026-11-23 首版（R73 派单 · 批 2 · 序 7）
//==============================================================================

(*------------------------------------------------------------------------------
 * 调用示例：fMR := FC_DL_MovingRangeCalc(fNewSample := x_i,
 *                                        fPrevSample := x_im1,
 *                                        bValid => bOk);
 * 注意：滑动窗历史驻留在上层 FB，本件只做相邻差值，两拍调用间无状态。
 * 组装说明：① 上层滑动窗管理件持有 x_(i−1) 并在下一拍回传 fPrevSample，
 *             本件零跨拍状态、可重入；
 *           ② 连续多拍极差进入 SPC 控制图判稳判据前，须校 bValid；
 *           ③ 本件输出单位与输入工程单位一致（差值不改单位）。
 *-----------------------------------------------------------------------------*)
FUNCTION FC_DL_MovingRangeCalc : LREAL
VAR_INPUT
    fNewSample  : LREAL;               // 本拍新样本 [工程单位随调用方] / New sample this scan [unit per caller]
    fPrevSample : LREAL;               // 上一拍样本 [工程单位随调用方] / Previous sample [unit per caller]
END_VAR
VAR_OUTPUT
    bValid      : BOOL;                // 结果有效标志，FALSE 时返回哨兵 0.0 / Result validity flag
END_VAR
VAR CONSTANT
    DL_MR_INF   : LREAL := 1.7976931348623157E308; // LREAL 幅值上限 / LREAL magnitude ceiling
    DL_MR_ZERO  : LREAL := 0.0;        // 无效哨兵返回值 / Sentinel return for invalid
END_VAR

// ---- 段 1｜出口默认值（纯函数无实例，无定时器/沿刷新义务）----
bValid := FALSE;                      // 缺省无效 / Invalid by default

// ---- 段 2｜输入防御：非有限值（NaN 自反判 + Inf 幅值判，R79）----
IF (fNewSample <> fNewSample) OR (ABS(fNewSample) > DL_MR_INF)
   OR (fPrevSample <> fPrevSample) OR (ABS(fPrevSample) > DL_MR_INF) THEN
    FC_DL_MovingRangeCalc := DL_MR_ZERO; // 无效输入：哨兵零返回，不进入运算 / Invalid input, sentinel zero return
    RETURN;                            // 结构早退 / early exit
END_IF

// ---- 段 3｜极差主体：MR = |x_i − x_(i−1)|，恒非负 ----
FC_DL_MovingRangeCalc := ABS(fNewSample - fPrevSample); // 滑动极差 / Moving range
bValid := TRUE;                       // 全部防御通过：结果有效 / Result valid
END_FUNCTION

(* ---- FC_DL_MultiPointLinear.st ---- *)
(*==============================================================================
 * 组件名称 (Component)  : FC_DL_MultiPointLinear
 * 所属子库 (Sublibrary) : DL_MathData
 * 当前版本 (Version)    : 1.0.0
 * 兼容性   (Platform)   : CODESYS 3.5 / TwinCAT 3 / 汇川 InoProShop / Machine Expert
 *                         仅依赖 Standard.library（ABS），全 LREAL 运算，无状态
 * 功能描述 (Function)   : N 段折线查表线性插值（N = 2..16）。用于热电偶、异形卧式罐液位、
 *                         流量计非线性修正、阀门特性补偿等"两点直线表达不了"的标定场景。
 *                         二分查找定位区间（O(log2 N)），输出命中段号与外推/钳位标志；
 *                         区间外默认钳位，显式关闭钳位才做端点段线性外推。
 *
 * 【失真与语义披露 / Distortion disclosure】
 *   1) 表非法（X 非严格递增）时整表作废，返回 afY[0]。这是刻意的"整体拒绝"：
 *      重复折点是除零的根因，若做"跳过坏点"的局部修补，会在现场产生一段斜率错误
 *      却看起来正常的插值，比直接报错危险得多。
 *   2) 非法表返回 afY[0] 而不是 0.0：0.0 在液位/温度场景会被当成真实测量值参与联锁，
 *      afY[0] 至少落在量程内，异常时工艺侧只会看到"读数不动"而不会看到"读数归零"。
 *   3) 外推在传感器断线时会把 0 mA 放大成负温度，因此默认钳位。要用外推必须显式
 *      把 bClamp 置 FALSE，并在设计文件中留档理由。
 *   4) 本函数不检测 NaN/Inf：IEC 61131-3 无标准判据，强行判断会引入编译器方言。
 *
 * 开源溯源 (Origin)     : 原创实现（参考西门子 LGF 定标族的"折线表 = X/Y 双数组 + 点数"
 *                         接口形态与 LBP 折线转换的粒度，clean-room 编写，未复制任何源码）
 * 依赖     (Depends)    : 无 DL_ 内部依赖；Standard.library: ABS
 * 红线自检 (Redline)    : R1 ✓ 零全局变量表与外部变量引用 ｜ R2 ✓ 零物理 IO 地址直写
 *                         R3 ✓ 纯 IEC 61131-3（无指针、无厂商私有符号）
 *                         R4 ✓ 点数钳位 + 单调性全校验 + 二分防死锁 + 段宽二次判零
 *                         R5 ✓ 全变量中英双语同行注释 ｜ R6 N/A（无状态机）｜ R7 N/A（无实例调用）
 * 修订历史 (Revision)   :
 *   2026-11-14  v1.0.0  首版入库（Phase 1 收口批次 · R3）
 *============================================================================*)
FUNCTION FC_DL_MultiPointLinear : LREAL
VAR_IN_OUT
    afX : ARRAY[0..15] OF LREAL;          // 折点自变量表，须严格递增（上限 16 点）/ Breakpoint X table, strictly increasing, max 16
    afY : ARRAY[0..15] OF LREAL;          // 折点因变量表 [EU]（上限 16 点）/ Breakpoint Y table [EU], max 16
END_VAR
VAR_INPUT
    fIn    : LREAL;                       // 输入值 [EU] / Input value [EU]
    nCount : INT;                         // 有效折点数，合法域 2..16 / Valid point count, 2..16
    bClamp : BOOL := TRUE;                // TRUE = 区间外钳位，FALSE = 线性外推 / TRUE = clamp, FALSE = extrapolate
END_VAR
VAR_OUTPUT
    nSegment      : INT;                  // 命中段号 0..nCount-2，-1 = 无效 / Segment index, -1 = invalid
    bExtrapolated : BOOL;                 // 本次结果来自外推 / Result comes from extrapolation
    bClamped      : BOOL;                 // 本次结果被钳位 / Result was clamped
    uErrorId      : UDINT;                // 故障码，0 = 无故障 / Error code, 0 = no error
END_VAR
VAR
    nLo      : INT;                       // 二分下界 / Binary search low bound
    nHi      : INT;                       // 二分上界 / Binary search high bound
    nMid     : INT;                       // 二分中点 / Binary search middle
    nGuard   : INT;                       // 二分防死锁计数器 / Binary search guard counter
    nIdx     : INT;                       // 单调性校验索引 / Monotonicity check index
    fX0      : LREAL;                     // 段左折点 X / Left breakpoint X
    fX1      : LREAL;                     // 段右折点 X / Right breakpoint X
    fY0      : LREAL;                     // 段左折点 Y [EU] / Left breakpoint Y [EU]
    fY1      : LREAL;                     // 段右折点 Y [EU] / Right breakpoint Y [EU]
    fSpan    : LREAL;                     // 段宽 fX1 - fX0 / Segment span
    fRatio   : LREAL;                     // 段内归一化位置，可越 0..1（外推时）/ Normalised position, may leave 0..1
    bTableOk : BOOL;                      // 表合法性标志 / Table validity flag
    bSearchOk: BOOL;                      // 二分收敛标志 / Binary search convergence flag
END_VAR
VAR CONSTANT
    DL_MPL_PTS_MIN : INT   := 2;          // 最少折点数 / Minimum point count
    DL_MPL_PTS_MAX : INT   := 16;         // 最多折点数，等于数组维度 / Maximum point count, equals the array size
    DL_MPL_EPS     : LREAL := 1.0E-9;     // 折点严格递增容差 / Strict-increase tolerance
    DL_MPL_GUARD   : INT   := 8;          // 二分最大迭代次数，log2(16)=4 留一倍余 / Max binary iterations
END_VAR

(*------------------------------------------------------------------------------
 * 段 1｜安全预置：返回值先落到表首值，异常路径不引入"0 值"这种伪测量
 *      Safe preset: default to the first table value, never to a fake zero
 *-----------------------------------------------------------------------------*)
FC_DL_MultiPointLinear := afY[0];
nSegment               := -1;
bExtrapolated          := FALSE;
bClamped               := FALSE;
uErrorId               := 16#0000_0000;
bTableOk               := TRUE;
bSearchOk              := TRUE;

(*------------------------------------------------------------------------------
 * 段 2｜点数校验（边界 B6）：先卡死点数，后面所有循环与索引才有定义域
 *      Point-count check first, so every later loop and index is well defined
 *-----------------------------------------------------------------------------*)
IF (nCount < DL_MPL_PTS_MIN) OR (nCount > DL_MPL_PTS_MAX) THEN
    uErrorId := 16#0001_0001;
    RETURN;
END_IF

(*------------------------------------------------------------------------------
 * 段 3｜单调性全校验（边界 B1）：整表拒绝，不做局部修补
 *      Whole-table monotonicity check: reject the whole table, never patch a bad point
 *-----------------------------------------------------------------------------*)
FOR nIdx := 1 TO (nCount - 1) DO
    IF (afX[nIdx] - afX[nIdx - 1]) <= DL_MPL_EPS THEN
        bTableOk := FALSE;
    END_IF
END_FOR

IF NOT bTableOk THEN
    uErrorId := 16#0002_000B;
    RETURN;
END_IF

(*------------------------------------------------------------------------------
 * 段 4｜区间外处理（边界 B3）：钳位优先，外推必须显式关闭
 *      Out-of-range handling: clamping wins, extrapolation must be opted in
 *-----------------------------------------------------------------------------*)
IF (fIn < afX[0]) AND bClamp THEN
    FC_DL_MultiPointLinear := afY[0];
    nSegment               := 0;
    bClamped               := TRUE;
    RETURN;
END_IF

IF (fIn > afX[nCount - 1]) AND bClamp THEN
    FC_DL_MultiPointLinear := afY[nCount - 1];
    nSegment               := (nCount - 2);
    bClamped               := TRUE;
    RETURN;
END_IF

IF (fIn < afX[0]) OR (fIn > afX[nCount - 1]) THEN
    bExtrapolated := TRUE;
END_IF

(*------------------------------------------------------------------------------
 * 段 5｜二分定位（边界 R4）：WHILE 必带防死锁计数器，超限强制收敛
 *      Binary search with a mandatory guard: over the limit it force-converges
 *      收敛判据是 nHi - nLo > 1，循环退出时必然 nLo ∈ 0..nCount-2，段号天然合法
 *-----------------------------------------------------------------------------*)
nLo := 0;
nHi := (nCount - 1);
nGuard := 0;

WHILE (nHi - nLo) > 1 DO

    nGuard := nGuard + 1;

    IF nGuard > DL_MPL_GUARD THEN
        (* 理论上不可达（4 次足够），纯防御：强制收敛并报保护触发 *)
        (* Unreachable in theory, pure defence: force convergence and report *)
        bSearchOk := FALSE;
        nHi       := (nLo + 1);
    ELSE
        nMid := (nLo + nHi) / 2;
        IF fIn >= afX[nMid] THEN
            nLo := nMid;
        ELSE
            nHi := nMid;
        END_IF
    END_IF

END_WHILE

IF NOT bSearchOk THEN
    uErrorId := 16#0001_0004;
END_IF

nSegment := nLo;

(*------------------------------------------------------------------------------
 * 段 6｜段内线性插值（边界 B4）：单调性已保证段宽 > EPS，这里仍再判一次
 *      Segment interpolation: the span is checked again, the table may be rewritten outside
 *      fIn 恰好等于折点时 fRatio = 1.0，结果等于该折点 Y，无跳变（边界 B5）
 *-----------------------------------------------------------------------------*)
fX0 := afX[nLo];
fX1 := afX[nLo + 1];
fY0 := afY[nLo];
fY1 := afY[nLo + 1];
fSpan := fX1 - fX0;

IF ABS(fSpan) > DL_MPL_EPS THEN
    fRatio := (fIn - fX0) / fSpan;
    FC_DL_MultiPointLinear := fY0 + fRatio * (fY1 - fY0);
ELSE
    (* 表在两次校验之间被外部改写：退回左折点值并报表非法 *)
    (* The table was rewritten between the checks: fall back to the left point *)
    FC_DL_MultiPointLinear := fY0;
    nSegment               := -1;
    uErrorId               := 16#0002_000B;
END_IF
END_FUNCTION

(* ---- FC_DL_Mux2Ex.st ---- *)
(*
    FC_DL_Mux2Ex —— 2 通道多路选择泛型防御包装（REAL 域）
    ------------------------------------------------------------------
    分类      : DL_MathData / Sel
    前缀      : FC_DL_
    版本      : 1.0.0
    溯源      : IEC 61131-3 标准语义的道莅防御性实现
                （内部委托平台内建函数，外围统一错误码/钳位/双语文档；
                  未复制任何闭源厂商源码，参考实现仅限 MIT/Apache 许可）
    平台      : 纯 IEC 61131-3，CODESYS / TwinCAT / InoProShop 通用
    作者      : 道莅代码库 · PLC编程专家（R16）
    ------------------------------------------------------------------
    功能说明  : 2 通道多路选择：uK=0 选 fI0、uK=1 选 fI1，选择运算用比较与
                IF/ELSE 实现（IEC MUX 语义），不重实现任何数学内核；
                uK 超出 0~1 时防御性钳位至 1，置信息级 16#0001_01D6（bError=FALSE、bValid=TRUE）；
                钳位方向：选择子越界单侧钳至上界 1；
                选中通道非有限（NaN 或 ±INF）判为故障级 16#0001_02AF，返回 0.0 且 bValid=FALSE；
                ±INF 采用平台安全幅值比较判定（阈值高于 REAL 最大有限值 3.402823E38），NaN 用自不等判定。
    错误码    : 16#0001_01D6 选择子 uK 越界，已钳位至 1——信息级，正常防御
                16#0001_02AF 选中通道非有限（NaN 或 ±INF）——故障级，返回 0.0
                16#0001_01D7 预留禁用（信息级，不得挪用）
                16#0001_02B0 预留禁用（故障级，不得挪用）
                16#0001_02B1 预留禁用（故障级，不得挪用）
    状态机    : R6 标注 N/A —— 本组件为纯函数无顺序状态机，无 CASE 可写，非法状态不可能出现，故以本节说明替代 ELSE 兜底
    修订记录  : 2026-11-16 v1.0.0 首次入库（R16）
*)
FUNCTION FC_DL_Mux2Ex : REAL
VAR_INPUT
    uK  : USINT; // 选择子 [通道号]，0~1，越界钳 1 / selector index [channel], 0~1, clamped to 1
    fI0 : REAL;  // 通道 0 输入 [无量纲] / channel 0 input
    fI1 : REAL;  // 通道 1 输入 [无量纲] / channel 1 input
END_VAR
VAR_OUTPUT
    eErr   : UDINT; // 错误码，0=正常 / error id, 0=ok
    bError : BOOL;  // 是否出错，eErr 非 0 时为 TRUE / error flag, TRUE when eErr is nonzero
    bValid : BOOL;  // 输出是否有效可用 / output valid flag
END_VAR
VAR CONSTANT
    DL_MUX2_CH_MAX    : USINT := 1;     // 通道选择子上界 [通道号] / selector index upper bound
    DL_REAL_INF_GUARD : LREAL := 4.0E38; // REAL 域 ±INF 判定阈值，高于 REAL 最大有限值 3.402823E38 [无量纲] / REAL +/-INF guard above max finite REAL 3.402823E38
END_VAR
VAR
    uIdx      : USINT; // 钳位后的本地选择子 [通道号] / clamped local selector index
    fSel      : REAL;  // 选中通道值 [无量纲] / selected channel value
    bSelBad   : BOOL;  // 选中通道非有限判定结果 / non-finite detection result of selected channel
END_VAR

// 段 1｜返回值与错误状态预置 / segment 1, preset return value and error status
FC_DL_Mux2Ex := 0.0; // 故障缺省返回 0 [无量纲] / fault default returns 0
eErr   := 0;     // 预置无错误 / preset no error
bError := FALSE; // 预置无故障 / preset no fault
bValid := FALSE; // 预置无效，通过防御闸后置位 / preset invalid, set TRUE after guard passes

// 段 2｜选择子越界钳位与通道选择 / segment 2, selector out-of-range clamp and channel selection
IF uK > DL_MUX2_CH_MAX THEN
    uIdx := DL_MUX2_CH_MAX; // 越界钳位至上界 1 / out-of-range clamped to upper bound 1
    eErr := 16#0001_01D6;   // 信息级：选择子越界已钳位 / info level: selector out of range, clamped
ELSE
    uIdx := uK; // 选择子在域内直通 / in-range selector passes through
END_IF
IF uIdx = 0 THEN
    fSel := fI0; // 通道 0 选中 / channel 0 selected
ELSE
    fSel := fI1; // 通道 1 选中（钳位后 uIdx 仅剩 0 或 1） / channel 1 selected (uIdx is only 0 or 1 after clamp)
END_IF

// 段 3｜选中通道防御闸与输出（末段） / segment 3, selected channel guard and output (final)
bSelBad := (fSel <> fSel) OR (fSel > DL_REAL_INF_GUARD) OR (fSel < -DL_REAL_INF_GUARD); // 选中通道非有限判定（NaN 自不等 + 安全幅值判 ±INF） [无量纲] / selected channel non-finite check (NaN by self-inequality, +/-INF by safe magnitude)
IF bSelBad THEN
    FC_DL_Mux2Ex := 0.0;      // 故障级返回 0 [无量纲] / fault level returns 0
    eErr   := 16#0001_02AF;   // 选中通道非有限故障码 / selected channel non-finite fault id
    bError := TRUE;           // 置故障标志 / set fault flag
    bValid := FALSE;          // 输出无效 / output invalid
    RETURN;                   // 立即返回 / immediate return
END_IF
bError := FALSE; // 信息级钳位不置故障，故障分支已提前返回 / info-level clamp never raises fault, fault branch has returned
bValid := TRUE;  // 选中通道输出有效可用 / selected channel output is valid
FC_DL_Mux2Ex := fSel; // 输出选中通道值 [无量纲] / output selected channel value
END_FUNCTION

(* ---- FC_DL_Mux4Ex.st ---- *)
(*
    FC_DL_Mux4Ex —— 4 通道多路选择泛型防御包装（REAL 域）
    ------------------------------------------------------------------
    分类      : DL_MathData / Sel
    前缀      : FC_DL_
    版本      : 1.0.0
    溯源      : IEC 61131-3 标准语义的道莅防御性实现
                （内部委托平台内建函数，外围统一错误码/钳位/双语文档；
                  未复制任何闭源厂商源码，参考实现仅限 MIT/Apache 许可）
    平台      : 纯 IEC 61131-3，CODESYS / TwinCAT / InoProShop 通用
    作者      : 道莅代码库 · PLC编程专家（R16）
    ------------------------------------------------------------------
    功能说明  : 4 通道多路选择：uK=0~3 分别选 fI0~fI3，选择运算用比较与
                IF/ELSIF 链实现（IEC MUX 语义），不重实现任何数学内核；
                uK 超出 0~3 时防御性钳位至 3，置信息级 16#0001_01D8（bError=FALSE、bValid=TRUE）；
                钳位方向：选择子越界单侧钳至上界 3；
                选中通道非有限（NaN 或 ±INF）判为故障级 16#0001_02B2，返回 0.0 且 bValid=FALSE；
                ±INF 采用平台安全幅值比较判定（阈值高于 REAL 最大有限值 3.402823E38），NaN 用自不等判定。
    错误码    : 16#0001_01D8 选择子 uK 越界，已钳位至 3——信息级，正常防御
                16#0001_02B2 选中通道非有限（NaN 或 ±INF）——故障级，返回 0.0
                16#0001_01D9 预留禁用（信息级，不得挪用）
                16#0001_02B3 预留禁用（故障级，不得挪用）
                16#0001_02B4 预留禁用（故障级，不得挪用）
    状态机    : R6 标注 N/A —— 本组件为纯函数无顺序状态机，无 CASE 可写，非法状态不可能出现，故以本节说明替代 ELSE 兜底
    修订记录  : 2026-11-16 v1.0.0 首次入库（R16）
*)
FUNCTION FC_DL_Mux4Ex : REAL
VAR_INPUT
    uK  : USINT; // 选择子 [通道号]，0~3，越界钳 3 / selector index [channel], 0~3, clamped to 3
    fI0 : REAL;  // 通道 0 输入 [无量纲] / channel 0 input
    fI1 : REAL;  // 通道 1 输入 [无量纲] / channel 1 input
    fI2 : REAL;  // 通道 2 输入 [无量纲] / channel 2 input
    fI3 : REAL;  // 通道 3 输入 [无量纲] / channel 3 input
END_VAR
VAR_OUTPUT
    eErr   : UDINT; // 错误码，0=正常 / error id, 0=ok
    bError : BOOL;  // 是否出错，eErr 非 0 时为 TRUE / error flag, TRUE when eErr is nonzero
    bValid : BOOL;  // 输出是否有效可用 / output valid flag
END_VAR
VAR CONSTANT
    DL_MUX4_CH_MAX    : USINT := 3;     // 通道选择子上界 [通道号] / selector index upper bound
    DL_REAL_INF_GUARD : LREAL := 4.0E38; // REAL 域 ±INF 判定阈值，高于 REAL 最大有限值 3.402823E38 [无量纲] / REAL +/-INF guard above max finite REAL 3.402823E38
END_VAR
VAR
    uIdx    : USINT; // 钳位后的本地选择子 [通道号] / clamped local selector index
    fSel    : REAL;  // 选中通道值 [无量纲] / selected channel value
    bSelBad : BOOL;  // 选中通道非有限判定结果 / non-finite detection result of selected channel
END_VAR

// 段 1｜返回值与错误状态预置 / segment 1, preset return value and error status
FC_DL_Mux4Ex := 0.0; // 故障缺省返回 0 [无量纲] / fault default returns 0
eErr   := 0;     // 预置无错误 / preset no error
bError := FALSE; // 预置无故障 / preset no fault
bValid := FALSE; // 预置无效，通过防御闸后置位 / preset invalid, set TRUE after guard passes

// 段 2｜选择子越界钳位与通道选择（IF/ELSIF 链实现 MUX 语义） / segment 2, selector out-of-range clamp and channel selection via IF/ELSIF chain (MUX semantics)
IF uK > DL_MUX4_CH_MAX THEN
    uIdx := DL_MUX4_CH_MAX; // 越界钳位至上界 3 / out-of-range clamped to upper bound 3
    eErr := 16#0001_01D8;   // 信息级：选择子越界已钳位 / info level: selector out of range, clamped
ELSE
    uIdx := uK; // 选择子在域内直通 / in-range selector passes through
END_IF
IF uIdx = 0 THEN
    fSel := fI0; // 通道 0 选中 / channel 0 selected
ELSIF uIdx = 1 THEN
    fSel := fI1; // 通道 1 选中 / channel 1 selected
ELSIF uIdx = 2 THEN
    fSel := fI2; // 通道 2 选中 / channel 2 selected
ELSE
    fSel := fI3; // 通道 3 选中（钳位后 uIdx 仅剩 0~3，此分支覆盖 uIdx=3） / channel 3 selected (uIdx is 0~3 after clamp, this branch covers uIdx=3)
END_IF

// 段 3｜选中通道防御闸与输出（末段） / segment 3, selected channel guard and output (final)
bSelBad := (fSel <> fSel) OR (fSel > DL_REAL_INF_GUARD) OR (fSel < -DL_REAL_INF_GUARD); // 选中通道非有限判定（NaN 自不等 + 安全幅值判 ±INF） [无量纲] / selected channel non-finite check (NaN by self-inequality, +/-INF by safe magnitude)
IF bSelBad THEN
    FC_DL_Mux4Ex := 0.0;      // 故障级返回 0 [无量纲] / fault level returns 0
    eErr   := 16#0001_02B2;   // 选中通道非有限故障码 / selected channel non-finite fault id
    bError := TRUE;           // 置故障标志 / set fault flag
    bValid := FALSE;          // 输出无效 / output invalid
    RETURN;                   // 立即返回 / immediate return
END_IF
bError := FALSE; // 信息级钳位不置故障，故障分支已提前返回 / info-level clamp never raises fault, fault branch has returned
bValid := TRUE;  // 选中通道输出有效可用 / selected channel output is valid
FC_DL_Mux4Ex := fSel; // 输出选中通道值 [无量纲] / output selected channel value
END_FUNCTION

(* ---- FC_DL_MuxIntEx.st ---- *)
(*
    FC_DL_MuxIntEx —— MUX 八路选择防御包装（INT 域）
    ------------------------------------------------------------------
    分类      : DL_MathData / Mux
    前缀      : FC_DL_
    版本      : 1.0.0
    溯源      : IEC 61131-3 标准语义的道莅防御性实现
                （内部委托 MUX 内建选择语义，外围统一错误码/钳位/双语文档；
                  未复制任何闭源厂商源码，参考实现仅限 MIT/Apache 许可）
    平台      : 纯 IEC 61131-3，CODESYS / TwinCAT / InoProShop 通用
    作者      : 道莅代码库 · PLC编程专家（R40）
    ------------------------------------------------------------------
    功能说明  : 八路 INT 选择器：按 uSel 选择 nIn0 至 nIn7 之一输出（0 基选择）；
                部分平台对 MUX 内建越路数选择的返回值未定义（有的返回 0、有的
                返回末路、有的触发异常），本件把越界行为显式化为钳位防御；
                选择值越路数时钳边界输出：uSel < 0 钳至通道 0，置信息级
                16#0001_0497；uSel > 7 钳至通道 7，置信息级 16#0001_0498；
                选择主体用 IF/ELSIF 链实现（IEC MUX 语义，不重实现选择内核），
                钳位保证选择值恒落在 [0, 7] 内，链分支全覆盖；
                链尾 ELSE 为理论不可达兜底（nSelC 已钳 [0, 7]，R128 口径：
                ELSE 只兜非法值）——命中时按选择下越界处置：钳回通道 0 并复用
                16#0001_0497（R90 复用不新占码位）；
                信息级码属正常防御：bError=FALSE、bValid=TRUE，输出钳位后防御值。
    错误码    : 16#0001_0497 选择值下越界（uSel < 0），已钳至通道 0——信息级，正常防御
                16#0001_0498 选择值上越界（uSel > 7），已钳至通道 7——信息级，正常防御
                （R90 反证句：下越界与上越界两场景均无法由返回值观测——钳位后输出
                  为合法通道值且 bValid=TRUE 与域内选择组合相同，若不占码则现场无法
                  还原「选错路」方向，故两侧各占一码）
    状态机    : R6 标注 N/A —— 本组件为纯函数无顺序状态机，无 ENUM 状态可写，
                选择链 ELSE 兜底已在功能说明段声明
    修订记录  : 2026-11-19 v1.0.0 首次入库（R40 · 批 3 · T0 快车道）
*)
FUNCTION FC_DL_MuxIntEx : INT
VAR_INPUT
    uSel : INT; // 选择值（0 基），越界时钳至边界通道 ｜ selector (0-based), clamped to a boundary channel when out of range
    nIn0 : INT; // 通道 0 输入 [无量纲] ｜ channel 0 input
    nIn1 : INT; // 通道 1 输入 [无量纲] ｜ channel 1 input
    nIn2 : INT; // 通道 2 输入 [无量纲] ｜ channel 2 input
    nIn3 : INT; // 通道 3 输入 [无量纲] ｜ channel 3 input
    nIn4 : INT; // 通道 4 输入 [无量纲] ｜ channel 4 input
    nIn5 : INT; // 通道 5 输入 [无量纲] ｜ channel 5 input
    nIn6 : INT; // 通道 6 输入 [无量纲] ｜ channel 6 input
    nIn7 : INT; // 通道 7 输入 [无量纲] ｜ channel 7 input
END_VAR
VAR_OUTPUT
    eErr   : UDINT; // 错误码，0=正常，16#0001_04XX=信息级 ｜ error id, 0=ok, 16#0001_04XX=info level
    bError : BOOL;  // 是否出错，本件信息级防御不置 TRUE ｜ fault flag, never raised by the info-level defense of this unit
    bValid : BOOL;  // 输出是否有效可用 ｜ output valid flag
END_VAR
VAR CONSTANT
    DL_MUX_CH_MAX : INT := 7; // 最高通道号（八路 0 基）[通道] ｜ highest channel index (8 channels, 0-based)
END_VAR
VAR
    nSelC : INT; // 钳位后的有效选择值 [通道] ｜ clamped effective selector
END_VAR

// 段 1｜返回值与错误状态预置 ｜ segment 1, preset return value and error status
FC_DL_MuxIntEx := 0; // 故障缺省返回 0 [无量纲] ｜ fault default returns 0
eErr   := 0;     // 预置无错误 ｜ preset no error
bError := FALSE; // 预置无故障 ｜ preset no fault
bValid := FALSE; // 预置无效，通过防御闸后置位 ｜ preset invalid, set TRUE after guard passes
nSelC  := 0;     // 选择值清零 ｜ clear the selector

// 段 2｜选择值越界钳位 ｜ segment 2, selector out-of-range clamp
IF uSel < 0 THEN
    nSelC := 0;             // 下越界钳至通道 0 [通道] ｜ under-range clamp to channel 0
    eErr  := 16#0001_0497;  // 信息级：下越界已钳位 ｜ info level: under-range clamped
ELSIF uSel > DL_MUX_CH_MAX THEN
    nSelC := DL_MUX_CH_MAX; // 上越界钳至通道 7 [通道] ｜ over-range clamp to channel 7
    eErr  := 16#0001_0498;  // 信息级：上越界已钳位 ｜ info level: over-range clamped
ELSE
    nSelC := uSel;          // 域内选择值直通 [通道] ｜ in-domain selector pass-through
END_IF

// 段 3｜选择主体（IF/ELSIF 链，末段） ｜ segment 3, selection body (IF/ELSIF chain, final)
IF nSelC = 0 THEN
    FC_DL_MuxIntEx := nIn0; // 通道 0 输出 [无量纲] ｜ channel 0 output
ELSIF nSelC = 1 THEN
    FC_DL_MuxIntEx := nIn1; // 通道 1 输出 [无量纲] ｜ channel 1 output
ELSIF nSelC = 2 THEN
    FC_DL_MuxIntEx := nIn2; // 通道 2 输出 [无量纲] ｜ channel 2 output
ELSIF nSelC = 3 THEN
    FC_DL_MuxIntEx := nIn3; // 通道 3 输出 [无量纲] ｜ channel 3 output
ELSIF nSelC = 4 THEN
    FC_DL_MuxIntEx := nIn4; // 通道 4 输出 [无量纲] ｜ channel 4 output
ELSIF nSelC = 5 THEN
    FC_DL_MuxIntEx := nIn5; // 通道 5 输出 [无量纲] ｜ channel 5 output
ELSIF nSelC = 6 THEN
    FC_DL_MuxIntEx := nIn6; // 通道 6 输出 [无量纲] ｜ channel 6 output
ELSIF nSelC = 7 THEN
    FC_DL_MuxIntEx := nIn7; // 通道 7 输出 [无量纲] ｜ channel 7 output
ELSE
    // 理论不可达兜底（nSelC 已钳 [0, 7]）：按选择下越界处置，复用 0497 不新占码位（R90）
    FC_DL_MuxIntEx := nIn0; // 兜底输出通道 0 [无量纲] ｜ backstop output of channel 0
    eErr := 16#0001_0497;   // 复用下越界信息码 ｜ reuse the under-range info code
END_IF
bError := FALSE; // 信息级钳位不置故障 ｜ info-level clamp never raises fault
bValid := TRUE;  // 域内或钳位输出均有效可用 ｜ in-domain or clamped output is valid
END_FUNCTION

(* ---- FC_DL_NormTo01.st ---- *)
(*
  ==================================================================
  组件名 Component  : FC_DL_NormTo01
  分类   Category   : DL_MathData
  前缀   Naming     : FC_DL_ ｜ b/n/u/f 类型前缀制（R265）
  版本   Version    : 1.0.0
  功能   Purpose    : 值域线性归一化至 0..1：fNorm = (fVal − fMin) /
                      (fMax − fMin)。反向域（fMax < fMin）与零域宽
                      （|fMax − fMin| < 容差，浮点容差判禁等号）双闸分
                      立；输入超 [fMin, fMax] 结果钳位至 0/1 并置信息码，
                      不静默。域宽为有限大数相减仍可能溢出 Inf，结果非
                      有限复核兜底。
  来源   Source     : t2-1-lgf-math（min-max 归一化为公开数学口径，
                      实现零源码复制）
  互引   Cross-ref  : FC_DL_Scaling（同族线性标定原子：其按工程量程
                      双点标定，本件为 0..1 归一口径属主）
  平台   Platform   : 纯 IEC 61131-3 四则 + ABS，三平台通用
  依赖   Depends    : 无 DL_ 内部依赖；无标准库
  红线   Redline    : R1 零全局/VAR_EXTERNAL/R2 零 %I/%Q/R3 纯 IEC 标准
                      R4 除零三闸（反向域/零域宽容差判/结果非有限复核）
                      + 钳位显式/R5 全变量双语同行注释/R6 纯函数无状态机
                      （CASE 不适用）/R7 无定时器与沿检测/R8 容差常量化
  错误码 Codes      : 01【失效级】反向域（fMax < fMin），返回 0
                      02【失效级】零域宽（|fMax − fMin| < 1E-9，浮点容差
                      判）或任一输入非有限或结果非有限，返回 0
                      03【信息级】超界钳位（fVal 出 [fMin,fMax]，结果钳
                      至 0 或 1，不置 bError）
  码位反证 Note     : 01/02 分立依据（R90）：01 在域序面（参数对调类组
                      态错）、02 在域宽/数值面（量程退化类组态错）可观测，
                      整定入口同但缺陷性质不同；03 信息级不置 bError，与
                      01/02 双通道可区分。
  验收   Acceptance : V1 fVal=fMin → 0 ｜ V2 fVal=fMax → 1 ｜ V3 中点 →
                      0.5 ｜ V4 fMax<fMin → 码 01 ｜ V5 fMax=fMin → 码 02
                      ｜ V6 超界 → 钳位 + 码 03（bValid=TRUE）
  变更   Revision   : 2026-11-22  v1.0.0  R67 首版（编码阶段批 2 序 3）
  ==================================================================
*)
FUNCTION FC_DL_NormTo01 : LREAL
VAR_INPUT
    fVal  : LREAL;  // 待归一值 [物理单位] / the value to normalize
    fMin  : LREAL;  // 域下界 [物理单位] / the domain lower bound
    fMax  : LREAL;  // 域上界 [物理单位] / the domain upper bound
END_VAR
VAR_OUTPUT
    bValid : BOOL;  // 归一值可用标志（钳位仍为 TRUE，头注 V6）[-] / the normalized value usable flag
    nErrId : UDINT; // 错误码，0=正常，01/02/03 见头注 [码] / the error code [code]
END_VAR
VAR
    fSpan  : LREAL; // 域宽工作寄存器 / the domain span working register
    fNorm  : LREAL; // 归一中间量工作寄存器 [-] / the normalized intermediate register
END_VAR
VAR CONSTANT
    N01_EPS     : LREAL := 1.0E-9;                 // 零域宽容差 [无量纲] / the zero span tolerance
    N01_FIN_MAX : LREAL := 1.7976931348623157E308; // LREAL 有限上限 / the finite LREAL limit
    N01_ERR_NONE : UDINT := 16#0000_0000;          // 无错误 [码] / no error [code]
    N01_ERR_REV  : UDINT := 16#0000_0001;          // 码 01：反向域 / code 01, reversed domain
    N01_ERR_ZSP  : UDINT := 16#0000_0002;          // 码 02：零域宽/非有限 / code 02, zero span or non finite
    N01_ERR_CLP  : UDINT := 16#0000_0003;          // 码 03：超界钳位（信息级）/ code 03, clamped, info level
END_VAR

// 段 1｜输出预置 / segment 1, preset the outputs
FC_DL_NormTo01 := 0.0;        // 失效缺省返回 0 / fault default returns zero
bValid := FALSE;              // 预置不可用 / preset unusable
nErrId := N01_ERR_NONE;       // 预置无错误 / preset no error

// 段 2｜输入非有限闸（并入码 02，头注口径）/ segment 2, the input finite gate
IF (fVal <> fVal) OR (fMin <> fMin) OR (fMax <> fMax)
   OR (ABS(fVal) > N01_FIN_MAX) OR (ABS(fMin) > N01_FIN_MAX) OR (ABS(fMax) > N01_FIN_MAX) THEN
    nErrId := N01_ERR_ZSP;
    RETURN;
END_IF

// 段 3｜反向域闸（码 01）：域序面缺陷 / segment 3, the reversed domain gate
IF fMax < fMin THEN
    nErrId := N01_ERR_REV;
    RETURN;
END_IF

// 段 4｜零域宽闸（码 02）：浮点容差判，禁 = 判等，除法前置 / segment 4, the zero span gate
fSpan := fMax - fMin;                      // 域宽（有限差可能 Inf，段 6 复核）/ the span
IF (ABS(fSpan) < N01_EPS) OR (fSpan <> fSpan) THEN
    nErrId := N01_ERR_ZSP;
    RETURN;
END_IF

// 段 5｜归一与超界钳位（码 03 信息级，钳位显式不静默）/ segment 5, normalize and clamp
fNorm := (fVal - fMin) / fSpan;            // 分母 = fSpan，已闸 / the denominator gated
IF (fNorm <> fNorm) OR (ABS(fNorm) > N01_FIN_MAX) THEN
    nErrId := N01_ERR_ZSP;                 // 结果非有限复核兜底 / the result finiteness recheck
    RETURN;
END_IF
IF fNorm < 0.0 THEN                        // 超下界钳 0 / clamp below
    fNorm := 0.0;
    nErrId := N01_ERR_CLP;
ELSIF fNorm > 1.0 THEN                     // 超上界钳 1 / clamp above
    fNorm := 1.0;
    nErrId := N01_ERR_CLP;
END_IF

// 段 6｜出口 / segment 6, the exit
FC_DL_NormTo01 := fNorm;                   // 归一值 [-] / the normalized value
bValid := TRUE;                            // 可用（钳位仍可用，头注 V6）/ usable, clamped still usable
END_FUNCTION

(* ---- FC_DL_OscillationIndex.st ---- *)
(*
  FC_DL_OscillationIndex  —  回路振荡指数（过零率 x 幅值离散度归一合成）/ Loop oscillation index
  分类 Category : DL_MathData
  码位 Code     : 16#05_0_03
  版本 Version  : 1.0.0
  来源 Source   : t2-4-s7-motion — IEC 61131-3 标准语义的道莅防御性实现
  溯源 Origin   : clean-room 实现，过零率与幅值离散度公开统计语义，未复制任何源码行
                  （与 FC_DL_CpkIndex 严格分工：本件判「在抖」— 振荡行为；FC_DL_CpkIndex 判「偏离」— 规格符合度）
  功能 Function : 1) 等间隔采样窗去均值后统计越过 ±fDeadband 的过零次数，得过零频率 fZeroCrossRateHz；
                  2) 幅值离散度 = 去均值绝对偏差均值 / 去均值幅值均值（fAmpDispersion）；
                  3) 两判据各自归一化后取几何平均合成 fOscIndex（0~1 无量纲），越 fOscNormLimit 判 bOscillating。
  边界 Boundary : ① nWindowSize < 8 或超数组上界判码（防越界）；② fSampleDt <= 0 防除零判码；
                  ③ 幅值均值 < fAmpFloor 判静止段：fOscIndex := 0 且 bOscillating := FALSE（不判抖）；
                  ④ fDeadband < 0 取 ABS 并置信息码（不拒算）；
                  ⑤ 非有限样本（NaN/Inf）按非法处理：本窗口无效置码，不输出指数；
                  ⑥ 解除式自证：bOscillating 每调用重算，下一窗指数回落即自动解除（无锁存）。
  依赖 Depends  : 仅 Standard.library（ABS/SQRT/MIN/MAX）；参考对齐 FB_DL_SignalStatistics（已注册，仅命名体例）；
                  分工件 FC_DL_CpkIndex（已注册，判偏离，与本件互不替代）
  码表 Error codes（本件格 05_0_03，子码步进 +0x100）:
    16#0005_0103 信息级：fDeadband 为负，已取 ABS 继续计算
    16#0005_0203 故障级：组态非法（窗长 < 8 / 超数组上界 / fSampleDt <= 0 / 归一化满量程 <= 0）
    16#0005_0303 故障级：采样窗含非有限值（NaN/Inf），本窗无效

  修订历史 Revision :
    2026-11-18  v1.0.0  R38 首版
*)

FUNCTION FC_DL_OscillationIndex : BOOL
VAR_INPUT
    afSampleBuffer : ARRAY[0..255] OF REAL;   // 等间隔采样窗 [工程量] / Equally spaced sample window
    nWindowSize    : INT;                     // 有效窗长 [点]，域 8..256 / Valid window length
    fSampleDt      : REAL;                    // 采样间隔 [s]，域 > 0 / Sample interval
    fDeadband      : REAL;                    // 判抖死区 [工程量单位] / Jitter deadband in engineering units
    fAmpFloor      : REAL := 0.01;            // 幅值均值下限 [工程量单位]，低于判静止 / Amplitude mean floor
    fNormRateHz    : REAL := 5.0;             // 过零率归一化满量程 [Hz]，域 > 0 / Zero-cross rate full-scale for normalization
    fOscNormLimit  : REAL := 0.3;             // 振荡判定阈值 [无量纲 0..1] / Oscillation verdict threshold
END_VAR
VAR_OUTPUT
    fOscIndex      : REAL;                    // 振荡指数 [无量纲 0..1] / Oscillation index
    fZeroCrossRateHz : REAL;                  // 过零频率 [Hz] / Zero-cross rate
    fAmpDispersion : REAL;                    // 幅值离散度 [无量纲] / Amplitude dispersion
    bOscillating   : BOOL;                    // 振荡判定 / Oscillation verdict
    nErrId         : UDINT;                   // 事件码，0 = 无事件 / Event code, 0 = none
END_VAR
VAR
    rMean, rAbsDev, rAmpMean : LREAL;         // 均值/绝对偏差和/幅值均值 / Mean, abs-deviation sum, amplitude mean
    rCross, rWinTime         : LREAL;         // 过零计数/窗时长 / Crossing count, window duration
    rRateN, rDispN, rIdx     : LREAL;         // 归一化过零率/归一化离散度/合成指数 / Normalized rate, dispersion, composite
    rD                       : LREAL;         // 单样本临时量 / Per-sample scratch
    rDb                      : LREAL;         // 死区生效值（负值取 ABS）/ Effective deadband
    k                        : INT;           // 循环计数器 / Loop counter
END_VAR
VAR CONSTANT
    nMinWin   : INT   := 8;       // 最小窗长 [点] / Minimum window length
    nMaxWin   : INT   := 256;     // 数组上界 [点] / Array upper bound
    rFinLim   : LREAL := 1.0E30;  // 非有限值筛查幅值上限 / Non-finite screening cap
    rDispNorm : LREAL := 1.0;     // 离散度归一化满量程（std/mean 量纲） / Dispersion full-scale
END_VAR

(* —— 段 1：输出缺省与组态闸（纯函数，每调用重算） —— *)
fOscIndex := 0.0;  fZeroCrossRateHz := 0.0;  fAmpDispersion := 0.0;   // 输出缺省
bOscillating := FALSE;                                                // 缺省不判抖（安全侧）
nErrId := 16#0000_0000;                                               // 事件码缺省无事件
FC_DL_OscillationIndex := FALSE;                                      // 返回值缺省失败

rDb := LREAL(fDeadband);                                              // 死区暂存
IF rDb < 0.0 THEN
    rDb := -rDb;                                                      // 负死区取 ABS 继续算（规格强制）
    nErrId := 16#0005_0103;                                           // 信息级：死区为负已取 ABS
END_IF

IF (nWindowSize < nMinWin) OR (nWindowSize > nMaxWin)
   OR (LREAL(fSampleDt) <= 0.0) OR (LREAL(fNormRateHz) <= 0.0) THEN
    nErrId := 16#0005_0203;                                           // 故障级：组态非法（覆盖防除零两项）
    RETURN;                                                           // 不进入计算
END_IF

(* —— 段 2：去均值 + 非有限值筛查（NaN 用 x<>x 自反判定，Inf 用幅值上限兜） —— *)
FOR k := 0 TO (nWindowSize - 1) DO
    rD := LREAL(afSampleBuffer[k]);
    IF (rD <> rD) OR (ABS(rD) > rFinLim) THEN
        nErrId := 16#0005_0303;                                       // 故障级：本窗含非有限值
        RETURN;                                                       // 整窗无效，不输出指数
    END_IF
    rMean := rMean + rD;                                              // 均值累加
END_FOR
rMean := rMean / LREAL(nWindowSize);                                  // 窗均值（窗长已闸 >= 8）

(* —— 段 3：幅值均值与过零计数（越过 ±死区计一次完整摆动） —— *)
FOR k := 0 TO (nWindowSize - 1) DO
    rD := LREAL(afSampleBuffer[k]) - rMean;                           // 去均值
    rAbsDev := rAbsDev + ABS(rD);                                     // 绝对偏差累加
END_FOR
rAmpMean := rAbsDev / LREAL(nWindowSize);                             // 幅值均值（平均绝对偏差）

FOR k := 1 TO (nWindowSize - 1) DO
    IF ((afSampleBuffer[k - 1] - REAL(rMean) < -REAL(rDb)) AND (afSampleBuffer[k] - REAL(rMean) >= REAL(rDb)))
       OR ((afSampleBuffer[k - 1] - REAL(rMean) > REAL(rDb)) AND (afSampleBuffer[k] - REAL(rMean) <= REAL(rDb))) THEN
        rCross := rCross + 1.0;                                       // 由 -侧 越到 +侧（或反向）：计 1 次过零
    END_IF
END_FOR

(* —— 段 4：静止段短路（幅值均值低于下限不判抖） —— *)
IF rAmpMean < LREAL(fAmpFloor) THEN
    fOscIndex := 0.0;                                                 // 静止段：指数 0
    bOscillating := FALSE;                                            // 不判抖（规格强制）
    FC_DL_OscillationIndex := TRUE;                                   // 计算已有效执行
    RETURN;                                                           // 过零率/离散度维持 0 缺省
END_IF

(* —— 段 5：频率与离散度归一化合成（分母均已闸） —— *)
rWinTime := LREAL(nWindowSize - 1) * LREAL(fSampleDt);                // 窗时长 [s]（fSampleDt 已闸 > 0）
IF rWinTime > 0.0 THEN
    fZeroCrossRateHz := REAL(rCross / (2.0 * rWinTime));              // 每次完整摆动含 2 次过零 [Hz]
END_IF
fAmpDispersion := REAL(MIN(rAmpMean / rDispNorm, 1.0));               // 离散度归一化并钳 0..1
rRateN := MIN(fZeroCrossRateHz / fNormRateHz, 1.0);                   // 过零率归一化并钳 0..1
rIdx := SQRT(rRateN * LREAL(fAmpDispersion));                         // 几何平均合成
fOscIndex := REAL(MIN(MAX(rIdx, 0.0), 1.0));                          // 钳 0..1

(* —— 段 6：判定出口 —— *)
bOscillating := fOscIndex > fOscNormLimit;                            // 越阈值判抖（每调用重算，解除式自证）
FC_DL_OscillationIndex := TRUE;                                       // 计算有效

END_FUNCTION

(* ---- FC_DL_PeakToPeakCalc.st ---- *)
(*
    FC_DL_PeakToPeakCalc —— 峰峰值计算（窗口 max−min + 非有限剔除 + 量程百分比）
    ------------------------------------------------------------------
    分类      : DL_MathData / Math-Statistics
    前缀      : FC_DL_
    版本      : 1.0.0
    来源标签  : iec-std-wrapper（T0）
    溯源      : IEC 61131-3 标准语义的道莅防御性实现
                （纯比较逻辑，无内建数学内核依赖；未复制任何闭源厂商源码）
    平台      : 纯 IEC 61131-3，CODESYS / TwinCAT / InoProShop 通用
    分工声明  : 与存量 FC_DL_SearchMinMax / FB_DL_WindowExtremaStat 分工——
                SearchMinMax 返回极值对本身，WindowExtremaStat 为驻留滑窗族；
                本件为无状态数组窗口峰峰值单出口并附量程百分比口径。
    作者      : 道莅代码库 · PLC 编程专家（R57）
    ------------------------------------------------------------------
    功能说明  : 对输入数组前 nCount 个样本求峰峰值（max−min）。窗长钳位
                ≥1（单样本峰峰值 0，边界十四）；非有限样本不参与并计数；
                fSpan <= 0 时百分比出口置 0 并置无效标志（防除零）。
    错误码    : 0000 正常 / 16#0003_0003 窗长已钳位 / 16#0003_0004 有效样本为零 / 16#0003_0006 量程组态非法
    修订记录  : 2026-11-21 v1.0.0 首次入库（R57 批 3 · 序号 14）
*)
FUNCTION FC_DL_PeakToPeakCalc : LREAL
VAR_IN_OUT
    afData : ARRAY[0..4095] OF LREAL; // 样本数组 [工程单位]，前 nCount 个有效 / the sample array, the first nCount entries valid
END_VAR
VAR_INPUT
    nCount : DINT; // 样本数 [个]，钳位 ≥1 / the sample count, clamped to one or above
    fSpan  : LREAL := 100.0; // 量程（用于百分比出口）[工程单位]，域 大于零 / the span for the percent outlet, above zero
END_VAR
VAR_OUTPUT
    eErr      : UDINT; // 错误码，0 = 正常 / error code, zero is ok
    bError    : BOOL;  // 出错标志，eErr 非 0 时为真 / error flag, true when eErr is nonzero
    bValid    : BOOL;  // 结果是否为真实值，钳位/剔除降级时为假 / the result is the true value, false when degraded
    fPctOfSpan: LREAL; // 峰峰值占量程百分比 [百分比] / the peak to peak over the span [percent]
    nNanCnt   : UDINT; // 剔除的非有限样本数 [个] / the excluded non finite sample count
    bPctValid : BOOL;  // 百分比出口有效性（fSpan 非法时为假）[-] / the percent outlet validity
END_VAR
VAR
    nI     : DINT;  // 循环计数 [个] / the loop counter
    nUsed  : DINT;  // 实际参与样本数 [个] / the used sample count
    lrMax  : LREAL; // 窗口最大值 [工程单位] / the window maximum
    lrMin  : LREAL; // 窗口最小值 [工程单位] / the window minimum
    lrX    : LREAL; // 当前样本 [工程单位] / the current sample
    bFirst : BOOL;  // 首个有效样本标记 [-] / the first valid sample flag
END_VAR

// 段 1｜返回值与错误状态预置安全值（四段式第一段，R45）/ segment 1, preset the return and error states
FC_DL_PeakToPeakCalc := 0.0; // 返回值预置安全值 0.0 / preset the return to the safe zero
fPctOfSpan := 0.0; // 百分比预置 0 / preset the percent zero
eErr   := 16#0000_0000; // 错误码预置正常 / preset the code to ok
bError := FALSE; // 错误标志预置假 / preset the error flag false
bValid := TRUE; // 有效标志预置真 / preset the valid flag true
bPctValid := TRUE; // 百分比有效性预置真 / preset the percent validity true
nNanCnt := 0; // 剔除计数预置零 / preset the excluded count zero
bFirst := TRUE; // 首样本标记预置真 / preset the first flag true
nUsed := 0; // 参与样本数预置零（防函数局部量残值）/ preset the used count zero

// 段 2｜窗长钳位 ≥1（边界十四）/ segment 2, the window clamp to one or above
IF nCount < 1 THEN // 低于下界 / below the floor
    nCount := 1; // 钳到 1 / clamp to one
    eErr   := 16#0003_0003; // 信息级：窗长已钳位 / informational, the window clamped
    bError := TRUE; // 置错误标志 / raise the error flag
    bValid := FALSE; // 钳位口径非原始口径 / the clamped window is not the requested one
END_IF

// 段 3｜量程组态闸（防除零，边界十四）/ segment 3, the span config gate against division by zero
IF (fSpan <= 0.0) OR (fSpan <> fSpan) OR ((fSpan - fSpan) <> (fSpan - fSpan)) THEN // 量程非法或非有限 / an illegal or non finite span
    fPctValid := FALSE; // 百分比出口置无效 / the percent outlet void
    eErr      := 16#0003_0006; // 信息级：量程组态非法 / informational, an illegal span config
    bError    := TRUE; // 置错误标志 / raise the error flag
END_IF

// 段 4｜窗口极值扫描（非有限剔除）/ segment 4, the extrema scan with exclusion
FOR nI := 0 TO nCount - 1 DO // 有界循环（nCount 已钳 ≤4096）/ the bounded loop
    lrX := afData[nI]; // 取样本（索引已证在数组界内）/ take the sample
    IF (lrX = lrX) AND ((lrX - lrX) = (lrX - lrX)) THEN // 非有限双判据通过才参与 / only finite samples participate
        IF bFirst THEN // 首个有效样本直接设为极值 / the first valid sample seeds both extrema
            lrMax := lrX; // 最大值播种 / seed the maximum
            lrMin := lrX; // 最小值播种 / seed the minimum
            bFirst := FALSE; // 播种完成 / the seeding done
        ELSE // 非首样本比较更新 / the later samples compared
            IF lrX > lrMax THEN // 超最大 / above the maximum
                lrMax := lrX; // 更新最大 / update the maximum
            END_IF
            IF lrX < lrMin THEN // 低于最小 / below the minimum
                lrMin := lrX; // 更新最小 / update the minimum
            END_IF
        END_IF
        nUsed := nUsed + 1; // 参与计数推进 / advance the used count
    ELSE // 非有限样本剔除 / a non finite sample excluded
        nNanCnt := nNanCnt + 1; // 剔除计数推进 / advance the excluded count
    END_IF
END_FOR

// 段 5｜结果计算 / segment 5, the result
IF nUsed > 0 THEN // 有有效样本 / with valid samples
    FC_DL_PeakToPeakCalc := lrMax - lrMin; // 峰峰值（单样本恰为 0，边界十四）/ the peak to peak, zero for a single sample
    IF bPctValid THEN // 量程合法才算百分比 / the percent only with a legal span
        fPctOfSpan := FC_DL_PeakToPeakCalc / fSpan * 100.0; // 百分比（除子已证大于零）/ the percent with a proven divisor
    END_IF
ELSE // 全部剔除 / all excluded
    eErr   := 16#0003_0004; // 错误级：有效样本为零 / error grade, no valid sample
    bError := TRUE; // 置错误标志 / raise the error flag
    bValid := FALSE; // 输出不可用 / the output void
END_IF
END_FUNCTION

(* ---- FC_DL_PearsonCorrCalc.st ---- *)
(*
  ==================================================================
  组件名 Component  : FC_DL_PearsonCorrCalc
  分类   Category   : DL_MathData
  前缀   Naming     : FC_DL_ ｜ b/n/u/f/t/e/st 类型前缀制（R265）
  码位   Code ID    : 16#0001_065B / 065C / 065D（故障级）｜ 16#0001_065E（信息级）
  版本   Version    : 1.0.0
  复杂度 Complexity  : 中
  功能   Purpose    : 双通道皮尔逊相关系数 r ∈ [−1, 1]，测点交叉诊断基元
                      （同源传感器相关失效、通道接错线检测）。
  开源溯源 Origin    : 公开公式 clean-room，参考公开统计学教材的皮尔逊积矩相关
                      定义（分类与公式借鉴，零代码复制），本件实现、闸门与码位
                      100% 自有。
  许可证 License    : MIT
  参考   Reference  : IEC 61131-3:2013 §6.6 算术运算符；Pearson r = Sxy /
                      SQRT(Sxx×Syy) 公开统计定义
  平台   Platform   : 纯 IEC 61131-3（FOR / 四则 / SQRT），三平台通用
  依赖   Depends    : 仅 Standard.library（SQRT 属标准内建）
  分工声明 Split     : FB_DL_CrossCorrelationDelay 为互相关时延估计属主（求滞后
                      拍数）；FB_DL_SensorPairPlausibility 为偏差 / 漂移互校；
                      本件为归一化相关强度；三件互引（R216）。SQRT 原语经派单
                      规格明写授权（除子 SQRT(Sxx×Syy)），本件为相关系数属主。
  归属 Ownership     : 本件无 TYPE 声明；全部引脚为 IEC 标准原生类型。
  ------------------------------------------------------------------
  边界 Boundary     :
                      一 配对剔除口径（写死）：X 或 Y 任一为非有限则**整对剔除**
                         （非各自剔除）——相关系数定义在样本对上，拆对剔除会
                         引入伪相关；nPairs = 剔除后有效对数；
                      二 nPairs ≤ 2（相关系数无定义）→ 故障码 065C 早退；
                      三 常量通道退化：Sxx ≤ 0 或 Syy ≤ 0（单通道方差为零，
                         相关系数无定义）→ 故障码 065D 早退（禁除零）；
                         ABS(Sxx×Syy) < 1.0E-12 防下溢分支同码处置（两场景出口
                         同形：fCorr = 0、bValid = FALSE，R90 不另立）；
                      四 数值口径：单遍累加 Σx / Σy / Σx² / Σy² / Σxy 后按
                         定义式展开（nPairs ≥ 3 已证，除子安全）；
                      五 |r| > 1.0（浮点数值误差）→ 钳回 ±1 并置信息级 065E
                         （不置 bError，R285）；
                      六 结果复检非有限 → 三件套兜底（R258）；
                      七 纯函数：无记忆量、无定时器、无边沿实例，每调用重算；
                      八 无全局、无外部变量、无物理地址、无指针。
  错误码 Codes      :
    16#0001_065B【故障级】样本对数越域（nCount < 1 / > 256）
    16#0001_065C【故障级】有效样本对数 ≤ 2（相关系数无定义）
    16#0001_065D【故障级】常量通道退化（Sxx ≤ 0 或 Syy ≤ 0）或乘积下溢
                         （ABS(Sxx×Syy) < 1.0E-12）
    16#0001_065E【信息级】|r| > 1.0 浮点数值误差，已钳回 ±1（不置 bError）
  码位反证 Note     :
    065B / 065C / 065D 三码不可合并：三者出口 nPairs 互异（越域 nPairs = 0、
    对数不足 nPairs ∈ [1,2]、常量退化 nPairs ≥ 3），可由 nPairs 唯一还原场景
    （R90）；065D 合并「常量通道」与「乘积下溢」：两场景出口组合同形
    （fCorr = 0、nPairs ≥ 3、bValid = FALSE），按 R90 不另立。
  验收 Acceptance   :
    算法已证（脚本）：未跑 ｜ 编译器已证（三平台）：未跑
    V1 完全线性 y = 2x → r ≈ +1（|r| ≤ 1 断言）；V2 y = −x → r ≈ −1
    V3 独立随机 → |r| < 0.1；V4 X 常数 → 码 065D 早退
    V5 单样本 / 双样本 → 码 065C 早退；V6 X 含 1 个 NaN → 整对剔除，
       nPairs 量化断言；V7 nCount = 0 → 码 065B
  修订记录 Revision  :
    2026-11-21  v1.0.0  R63 首版（批 2 · 序号 5）
  ==================================================================
*)
FUNCTION FC_DL_PearsonCorrCalc : BOOL
VAR_IN_OUT
    afX : ARRAY[0..255] OF LREAL; // 通道 X 样本 [工程单位]，只读 / the channel X samples, read only
    afY : ARRAY[0..255] OF LREAL; // 通道 Y 样本 [工程单位]，只读 / the channel Y samples, read only
END_VAR
VAR_INPUT
    nCount  : DINT := 0; // 样本对数入参 [对]，合法域 1..256 / the pair count, legal from one to two hundred fifty six
END_VAR
VAR_OUTPUT
    fCorr   : LREAL := 0.0; // 相关系数 [−]，−1..1 / the correlation coefficient inside the unit interval
    nPairs  : DINT := 0;    // 有效样本对数 [对]（配对剔除后）/ the effective pair count after the paired drop
    bValid  : BOOL := FALSE; // 结果可用 [-] / the result usable flag
    eErr    : UDINT := 16#0000_0000; // 错误码，0 = 正常 / the error code, zero is ok
    bError  : BOOL := FALSE; // 故障标志（故障级码同拍置位，R45 配对）/ the fault flag raised with a fault level code
END_VAR
VAR
    aXVal     : ARRAY[0..255] OF LREAL; // 剔除后 X 有效副本 [工程单位] / the effective copy of channel X
    aYVal     : ARRAY[0..255] OF LREAL; // 剔除后 Y 有效副本 [工程单位] / the effective copy of channel Y
    k         : DINT := 0;    // 遍历索引 [下标] / the traversal index
    nCountUse : DINT := 0;    // 入参对数接管量 [对] / the raw input count holder
    fSx       : LREAL := 0.0; // Σx 累加量 [工程单位] / the sum of x
    fSy       : LREAL := 0.0; // Σy 累加量 [工程单位] / the sum of y
    fSxx      : LREAL := 0.0; // Σx² 累加量 [工程单位²] / the sum of x squared
    fSyy      : LREAL := 0.0; // Σy² 累加量 [工程单位²] / the sum of y squared
    fSxy      : LREAL := 0.0; // Σxy 累加量 [工程单位²] / the sum of the cross products
    fMx       : LREAL := 0.0; // X 均值 [工程单位] / the mean of x
    fMy       : LREAL := 0.0; // Y 均值 [工程单位] / the mean of y
    fDxx      : LREAL := 0.0; // 中心化离差平方和 Sxx [工程单位²] / the centered sum of squares of x
    fDyy      : LREAL := 0.0; // 中心化离差平方和 Syy [工程单位²] / the centered sum of squares of y
    fDxy      : LREAL := 0.0; // 中心化叉积和 Sxy [工程单位²] / the centered cross product sum
    fDen      : LREAL := 0.0; // 归一化除子 SQRT(Sxx×Syy) [工程单位²] / the normalization divisor
    fCorrUse  : LREAL := 0.0; // 相关系数工作副本 [−] / the working correlation copy
    nPairsUse : DINT := 0;    // 有效对数工作副本 [对] / the working pair count
END_VAR  // R64 结构补齐：VAR 段缺失的 END_VAR（门禁机械修复）
VAR CONSTANT
    DL_PCC_NMAX  : DINT := 256;       // 样本容量上界 [对]，与数组容量一致 / the capacity aligned with the arrays
    DL_PCC_MIN   : DINT := 3;         // 相关系数可定义最少对数 [对] / the minimum pair count for a defined correlation
    DL_PCC_ONE   : DINT := 1;         // 整型一常量 [对] / the integer one constant
    DL_PCC_ZERO  : DINT := 0;         // 整型零常量 [对] / the integer zero constant
    DL_PCC_DENMIN: LREAL := 1.0E-12;  // 除子防下溢门限 [工程单位⁴] / the divisor underflow threshold
    DL_PCC_ONE_R : LREAL := 1.0;      // 单位一常量 [−]（钳位界）[-] / the unit constant used as the clamp bound
END_VAR

// 段 1｜返回值与全部出口预置安全值（R45 四段式第一段）/ segment 1, the preset of the return and every outlet
FC_DL_PearsonCorrCalc := FALSE; // 返回值预置假 / preset the return false
fCorr := 0.0; // 相关系数预置零 [−] / preset the correlation zero
nPairs := DL_PCC_ZERO; // 有效对数预置零 [对] / preset the pair count zero
bValid := FALSE; // 可用标志预置假 / preset the validity false
eErr := 16#0000_0000; // 错误码预置正常 / preset the code to ok
bError := FALSE; // 故障标志预置假 / preset the error flag false
nCountUse := DL_PCC_ZERO; // 入参对数接管量预置零 [对] / preset the raw count holder zero
nPairsUse := DL_PCC_ZERO; // 有效对数工作副本预置零 [对] / preset the working pair count zero
fSx := 0.0; // Σx 预置零 [工程单位] / preset the sum of x zero
fSy := 0.0; // Σy 预置零 [工程单位] / preset the sum of y zero
fSxx := 0.0; // Σx² 预置零 [工程单位²] / preset the sum of x squared zero
fSyy := 0.0; // Σy² 预置零 [工程单位²] / preset the sum of y squared zero
fSxy := 0.0; // Σxy 预置零 [工程单位²] / preset the cross sum zero
fMx := 0.0; // X 均值预置零 [工程单位] / preset the mean of x zero
fMy := 0.0; // Y 均值预置零 [工程单位] / preset the mean of y zero
fDxx := 0.0; // Sxx 预置零 [工程单位²] / preset the centered sum of squares zero
fDyy := 0.0; // Syy 预置零 [工程单位²] / preset the centered sum of squares zero
fDxy := 0.0; // Sxy 预置零 [工程单位²] / preset the centered cross sum zero
fDen := 0.0; // 除子预置零 [工程单位²] / preset the divisor zero
fCorrUse := 0.0; // 相关系数工作副本预置零 [−] / preset the working correlation zero
k := DL_PCC_ZERO; // 索引预置零 / preset the index zero

// 段 2｜样本对数域闸（边界八，早退禁除零）/ segment 2, the pair count domain gate
nCountUse := nCount; // 入参对数接管 [对] / take the raw count
IF (nCountUse < DL_PCC_ONE) OR (nCountUse > DL_PCC_NMAX) THEN // 对数越域 / the count is out of the domain
    eErr := 16#0001_065B; // 故障级：样本对数越域 / fault grade, the pair count is out of the domain
    bError := TRUE; // 同拍置故障标志（R45 配对）/ raise the fault flag on the same scan
    bValid := FALSE; // 结果不可用 / the result is not usable
    RETURN; // 早退 / early return
END_IF

// 段 3｜配对剔除（边界一：任一通道非有限则整对剔除）/ segment 3, the paired drop
FOR k := DL_PCC_ZERO TO nCountUse - DL_PCC_ONE DO // 有界遍历（上界已证 ≤ 256）/ the bounded traversal with a proven ceiling
    IF ((afX[k] = afX[k]) AND ((afX[k] - afX[k]) = (afX[k] - afX[k]))
    AND (afY[k] = afY[k]) AND ((afY[k] - afY[k]) = (afY[k] - afY[k]))) THEN // 整对有限 / the whole pair is finite
        aXVal[nPairsUse] := afX[k]; // X 写入有效副本 [工程单位] / copy the x sample
        aYVal[nPairsUse] := afY[k]; // Y 写入有效副本 [工程单位] / copy the y sample
        nPairsUse := nPairsUse + DL_PCC_ONE; // 有效对数推进 [对] / advance the pair count
    END_IF // 任一通道非有限：整对丢弃（不拆对）/ either channel broken, the whole pair is dropped
END_FOR
nPairs := nPairsUse; // 有效对数出口 [对] / export the pair count
IF nPairsUse < DL_PCC_MIN THEN // 有效对数 ≤ 2：相关系数无定义（边界二）/ too few pairs for a defined correlation
    eErr := 16#0001_065C; // 故障级：有效样本对数不足 / fault grade, the effective pairs are too few
    bError := TRUE; // 同拍置故障标志（R45 配对）/ raise the fault flag on the same scan
    bValid := FALSE; // 结果不可用 / the result is not usable
    RETURN; // 早退，除子段不可达 / early return, the divisor segment is unreachable
END_IF

// 段 4｜单遍累加（nPairs ≥ 3 已证，除子安全，边界四）/ segment 4, the single pass accumulation
FOR k := DL_PCC_ZERO TO nPairsUse - DL_PCC_ONE DO // 有界遍历有效对 / the bounded traversal over the effective pairs
    fSx := fSx + aXVal[k]; // Σx 累加 [工程单位] / accumulate the sum of x
    fSy := fSy + aYVal[k]; // Σy 累加 [工程单位] / accumulate the sum of y
    fSxx := fSxx + (aXVal[k] * aXVal[k]); // Σx² 累加 [工程单位²] / accumulate the sum of squares
    fSyy := fSyy + (aYVal[k] * aYVal[k]); // Σy² 累加 [工程单位²] / accumulate the sum of squares
    fSxy := fSxy + (aXVal[k] * aYVal[k]); // Σxy 累加 [工程单位²] / accumulate the cross products
END_FOR
fMx := fSx / DINT_TO_LREAL(nPairsUse); // X 均值 [工程单位]，除子已证 ≥ 3 / the mean of x with the proven divisor
fMy := fSy / DINT_TO_LREAL(nPairsUse); // Y 均值 [工程单位] / the mean of y
fDxx := fSxx - (DINT_TO_LREAL(nPairsUse) * fMx * fMx); // Sxx = Σx² − n·mx² [工程单位²] / the centered sum of squares of x
fDyy := fSyy - (DINT_TO_LREAL(nPairsUse) * fMy * fMy); // Syy = Σy² − n·my² [工程单位²] / the centered sum of squares of y
fDxy := fSxy - (DINT_TO_LREAL(nPairsUse) * fMx * fMy); // Sxy = Σxy − n·mx·my [工程单位²] / the centered cross product sum

// 段 5｜常量通道退化与除子防下溢闸（边界三，禁除零）/ segment 5, the constant channel and the underflow gate
IF (fDxx <= 0.0) OR (fDyy <= 0.0) OR (ABS(fDxx * fDyy) < DL_PCC_DENMIN) THEN // 常量通道或乘积下溢 / a constant channel or an underflowing product
    fCorr := 0.0; // 兜底安全值 [−] / the bottom line safe value
    eErr := 16#0001_065D; // 故障级：常量通道退化 / fault grade, a constant channel degeneration
    bError := TRUE; // 同拍置故障标志（R45 配对）/ raise the fault flag on the same scan
    bValid := FALSE; // 结果不可用 / the result is not usable
    RETURN; // 早退，除法不可达 / early return, the division is unreachable
END_IF

// 段 6｜相关系数计算（除子已证 > 0 且 ≥ 下溢门限）/ segment 6, the correlation computation
fDen := SQRT(fDxx * fDyy); // 归一化除子 [工程单位²]，已证有限且非零 / the normalization divisor proven finite and nonzero
fCorrUse := fDxy / fDen; // 皮尔逊相关系数 [−] / the Pearson correlation coefficient

// 段 7｜|r| > 1 钳位（浮点数值误差，信息级 065E，不置 bError）/ segment 7, the unit interval clamp with an informational code
IF ABS(fCorrUse) > DL_PCC_ONE_R THEN // 数值误差越单位圆 / a numerical overshoot beyond the unit circle
    IF fCorrUse > 0.0 THEN // 正向越界 / a positive overshoot
        fCorrUse := DL_PCC_ONE_R; // 钳回 +1 [−] / clamp to plus one
    ELSE // 负向越界 / a negative overshoot
        fCorrUse := -DL_PCC_ONE_R; // 钳回 −1 [−] / clamp to minus one
    END_IF
    eErr := 16#0001_065E; // 信息级：|r| 越界已钳回（不置 bError，R285）/ informational, the coefficient was clamped
END_IF

// 段 8｜结果复检兜底（三件套，R258）/ segment 8, the result recheck with the three part fallback
IF (fCorrUse <> fCorrUse) OR ((fCorrUse - fCorrUse) <> (fCorrUse - fCorrUse)) THEN // 结果非有限（理论上不可达，防御保留）/ a non finite result, unreachable by theory, kept as a defence
    fCorr := 0.0; // 兜底安全值 [−] / the bottom line safe value
    eErr := 16#0001_065D; // 故障级：常量通道退化（同族一码，出口组合不可区分，R90）/ fault grade under the same family code
    bError := TRUE; // 置故障标志（R45 配对）/ raise the fault flag
    bValid := FALSE; // 结果不可用 / the result is not usable
    RETURN; // 早退 / early return
END_IF

// 段 9｜统一出口 / segment 9, the unified outlet
fCorr := fCorrUse; // 相关系数出口 [−] / the correlation outlet
bValid := TRUE; // 结果可用 / the result is usable
FC_DL_PearsonCorrCalc := TRUE; // 返回成功 / return success
END_FUNCTION
